(* IEC 61131-3 sources: TetherPLC/compat/tc2, 47 files *)

(* ---- tc2_math.st ---- *)
// Tc2_Math compatibility functions (TwinCAT 3 PLC Library Tc2_Math).
// Pure LREAL math; sources from docs/plc/plan/21-twincat-libraries.md §7.
// Limitation: TRUNC narrows through DINT, so |x| >= 2^31 loses precision
// (same bound as Beckhoff's 32-bit TRUNC-based implementations).

FUNCTION F_TruncL : LREAL
VAR_INPUT
    lr_in : LREAL;
END_VAR
    F_TruncL := DINT_TO_LREAL(TRUNC(lr_in));
END_FUNCTION

FUNCTION CEIL : LREAL
VAR_INPUT
    lr_in : LREAL;
END_VAR
VAR
    t : LREAL;
END_VAR
    t := F_TruncL(lr_in);
    IF lr_in > t THEN
        CEIL := t + 1.0;
    ELSE
        CEIL := t;
    END_IF;
END_FUNCTION

FUNCTION FLOOR : LREAL
VAR_INPUT
    lr_in : LREAL;
END_VAR
VAR
    t : LREAL;
END_VAR
    t := F_TruncL(lr_in);
    IF lr_in < t THEN
        FLOOR := t - 1.0;
    ELSE
        FLOOR := t;
    END_IF;
END_FUNCTION

FUNCTION FRAC : LREAL
VAR_INPUT
    lr_in : LREAL;
END_VAR
    FRAC := lr_in - F_TruncL(lr_in);
END_FUNCTION

FUNCTION LTRUNC : LREAL
VAR_INPUT
    lr_in : LREAL;
END_VAR
    LTRUNC := F_TruncL(lr_in);
END_FUNCTION

FUNCTION LMOD : LREAL
VAR_INPUT
    lr_Value : LREAL;
    lr_Arg   : LREAL;
END_VAR
    IF lr_Arg = 0.0 THEN
        LMOD := 0.0;
    ELSE
        LMOD := lr_Value - F_TruncL(lr_Value / lr_Arg) * lr_Arg;
    END_IF;
END_FUNCTION

FUNCTION MODABS : LREAL
VAR_INPUT
    lr_val : LREAL;
    lr_mod : LREAL;
END_VAR
VAR
    am : LREAL;
END_VAR
    am := ABS(lr_mod);
    IF am = 0.0 THEN
        MODABS := 0.0;
    ELSE
        MODABS := lr_val - FLOOR(lr_val / am) * am;
    END_IF;
END_FUNCTION

FUNCTION MODTURNS : DINT
VAR_INPUT
    lr_Value : LREAL;
    lr_Arg   : LREAL;
END_VAR
    IF lr_Arg = 0.0 THEN
        MODTURNS := 0;
    ELSE
        MODTURNS := TRUNC(lr_Value / lr_Arg);
    END_IF;
END_FUNCTION

FUNCTION F_GetVersionTcMath : UINT
VAR_INPUT
    nVersionElement : INT;
END_VAR
    F_GetVersionTcMath := 16#0100;
END_FUNCTION

(* ---- tc2_ncdrive.st ---- *)
// Tc2_NcDrive — NC-axis SoE/CoE drive blocks.
//
// The 20 function blocks of this library are provided by
// compat/tc2/tc2_mc2_drive.st: the NcDrive variants take
// NCTOPLC_AXIS_REF + sNetId where the MC2_Drive variants take
// AXIS_REF + NetId, and both flatten to the same UDINT axis handle
// (slave = Axis - 1) over FB_Soe/FB_MotionAxis.  Covered:
//   FB_SoEReset, FB_SoEWritePassword, FB_SoEExecuteCommand,
//   FB_SoEWriteCommandControl, FB_SoEReadCommandState,
//   FB_SoEReadDiagMessage, FB_SoEReadDiagNumber,
//   FB_SoEReadDiagNumberList, FB_SoEReadClassXDiag, FB_SoERead,
//   FB_SoEWrite, FB_SoEReadAmplifierTemperature,
//   FB_SoEReadMotorTemperature, FB_SoEReadDcBusCurrent,
//   FB_SoEReadDcBusVoltage, FB_CoERead, FB_CoEWrite,
//   FB_SoEAX5000ReadActMainVoltage, FB_SoEAX5000SetMotorCtrlWord,
//   FB_SoEAX5000FirmwareUpdate.
// Deviations (shared with Tc2_MC2_Drive): PVOID buffers flatten to
// scalar Value members, tTimeout is not modeled, bCompleteAccess is
// accepted but sub-index access is unsupported, and the AX5000
// firmware update records the request only.

// F_GetVersionTcNcDrive — library version.
FUNCTION F_GetVersionTcNcDrive : UDINT
F_GetVersionTcNcDrive := 16#0100;
END_FUNCTION

(* ---- tc2_standard_wide.st ---- *)
// Tc2_Standard wide-string functions (TwinCAT 3 PLC Library Tc2_Standard).
// W* signatures mirror IEC 61131-3 string functions; bodies delegate to the
// same builtins, which already accept WSTRING operands.
// Sources: docs/plc/plan/21-twincat-libraries.md §7.

FUNCTION WCONCAT : WSTRING
VAR_INPUT
    STR1 : WSTRING;
    STR2 : WSTRING;
END_VAR
    WCONCAT := CONCAT(STR1, STR2);
END_FUNCTION

FUNCTION WDELETE : WSTRING
VAR_INPUT
    STR1 : WSTRING;
    LEN  : INT;
    POS  : INT;
END_VAR
    WDELETE := DELETE(STR1, LEN, POS);
END_FUNCTION

FUNCTION WFIND : INT
VAR_INPUT
    STR1 : WSTRING;
    STR2 : WSTRING;
END_VAR
    WFIND := FIND(STR1, STR2);
END_FUNCTION

FUNCTION WINSERT : WSTRING
VAR_INPUT
    STR1 : WSTRING;
    STR2 : WSTRING;
    POS  : INT;
END_VAR
    WINSERT := INSERT(STR1, STR2, POS);
END_FUNCTION

FUNCTION WLEFT : WSTRING
VAR_INPUT
    STR  : WSTRING;
    SIZE : INT;
END_VAR
    WLEFT := LEFT(STR, SIZE);
END_FUNCTION

FUNCTION WLEN : INT
VAR_INPUT
    STR : WSTRING;
END_VAR
    WLEN := LEN(STR);
END_FUNCTION

FUNCTION WMID : WSTRING
VAR_INPUT
    STR  : WSTRING;
    LEN  : INT;
    POS  : INT;
END_VAR
    WMID := MID(STR, LEN, POS);
END_FUNCTION

FUNCTION WREPLACE : WSTRING
VAR_INPUT
    STR1 : WSTRING;
    STR2 : WSTRING;
    L    : INT;
    P    : INT;
END_VAR
    WREPLACE := REPLACE(STR1, STR2, L, P);
END_FUNCTION

FUNCTION WRIGHT : WSTRING
VAR_INPUT
    STR  : WSTRING;
    SIZE : INT;
END_VAR
    WRIGHT := RIGHT(STR, SIZE);
END_FUNCTION

(* ---- tc2_aes70.st ---- *)
// tc2_aes70.st — TwinCAT audio-control client surface (Tc3_AES70 /
// TF6301-ish shape) over the tplc-aes70 service + FB_Aes70 builtin.
//
// The PLC is the OCA client over OSCP TCP (AES70/Open Control
// Architecture): FB_Aes70Connect opens the TCP session on the OCA
// control port (default 65000); FB_Aes70Call carries an OcaCommand
// (targetONo + methodID + parameter bytes);
// FB_Aes70Receive polls for a pending OcaResponse each scan;
// Keepalive sends an OSCP heartbeat; Disconnect releases.
//
// Parameters and response payloads are raw bytes bounded
// STRING[255] — the caller composes/parses the OCA-serialized
// parameter set.  Notification subscriptions, the full OCA class
// catalog, and property/get-set shorthands are out of scope for
// this tranche.

// ---- FB_Aes70Connect: TCP session on the OCA control port ----
FUNCTION_BLOCK FB_Aes70Connect
VAR_INPUT
    Execute : BOOL;
    Host : STRING[63];
    Port : UDINT;
END_VAR
VAR_OUTPUT
    Done : BOOL;
    Busy : BOOL;
    Error : BOOL;
    ErrorID : UDINT;
    ConnectionHdl : UDINT;
END_VAR
VAR
    ch : FB_Aes70;
    exPrev : BOOL;
END_VAR
    Done := FALSE;
    Error := FALSE;
    ErrorID := 0;
    IF Execute AND NOT exPrev THEN
        ch.OP := 1;
        ch.HOST := Host;
        ch.PORT := Port;
        ch();
        IF ch.STATUS = 0 THEN
            Done := TRUE;
            ConnectionHdl := ch.HANDLE;
        ELSE
            Error := TRUE;
            ErrorID := ch.ERRID;
        END_IF;
    END_IF;
    exPrev := Execute;
    Busy := FALSE;
END_FUNCTION_BLOCK

// ---- FB_Aes70Disconnect: release the session ----
FUNCTION_BLOCK FB_Aes70Disconnect
VAR_INPUT
    Execute : BOOL;
    ConnectionHdl : UDINT;
END_VAR
VAR_OUTPUT
    Done : BOOL;
    Busy : BOOL;
    Error : BOOL;
    ErrorID : UDINT;
END_VAR
VAR
    ch : FB_Aes70;
    exPrev : BOOL;
END_VAR
    Done := FALSE;
    Error := FALSE;
    ErrorID := 0;
    IF Execute AND NOT exPrev THEN
        ch.OP := 2;
        ch.HANDLE := ConnectionHdl;
        ch();
        IF ch.STATUS = 0 THEN
            Done := TRUE;
        ELSE
            Error := TRUE;
            ErrorID := ch.ERRID;
        END_IF;
    END_IF;
    exPrev := Execute;
    Busy := FALSE;
END_FUNCTION_BLOCK

// ---- FB_Aes70Call: OcaCommand on an object ----
FUNCTION_BLOCK FB_Aes70Call
VAR_INPUT
    Execute : BOOL;
    ConnectionHdl : UDINT;
    TargetONo : UDINT;
    MethodID : UDINT;
    Params : STRING[255];
END_VAR
VAR_OUTPUT
    Done : BOOL;
    Error : BOOL;
    ErrorID : UDINT;
    RequestHdl : UDINT;
END_VAR
VAR
    ch : FB_Aes70;
    exPrev : BOOL;
END_VAR
    Done := FALSE;
    Error := FALSE;
    ErrorID := 0;
    IF Execute AND NOT exPrev THEN
        ch.OP := 4;
        ch.HANDLE := ConnectionHdl;
        ch.TARGET := TargetONo;
        ch.METH := MethodID;
        ch.PARAMS := Params;
        ch();
        IF ch.STATUS = 0 THEN
            Done := TRUE;
            RequestHdl := ch.HANDLE2;
        ELSE
            Error := TRUE;
            ErrorID := ch.ERRID;
        END_IF;
    END_IF;
    exPrev := Execute;
END_FUNCTION_BLOCK

// ---- FB_Aes70Keepalive: OSCP heartbeat ----
FUNCTION_BLOCK FB_Aes70Keepalive
VAR_INPUT
    Execute : BOOL;
    ConnectionHdl : UDINT;
END_VAR
VAR_OUTPUT
    Done : BOOL;
    Error : BOOL;
    ErrorID : UDINT;
END_VAR
VAR
    ch : FB_Aes70;
    exPrev : BOOL;
END_VAR
    Done := FALSE;
    Error := FALSE;
    ErrorID := 0;
    IF Execute AND NOT exPrev THEN
        ch.OP := 5;
        ch.HANDLE := ConnectionHdl;
        ch();
        IF ch.STATUS = 0 THEN
            Done := TRUE;
        ELSE
            Error := TRUE;
            ErrorID := ch.ERRID;
        END_IF;
    END_IF;
    exPrev := Execute;
END_FUNCTION_BLOCK

// ---- FB_Aes70Receive: poll for a pending OcaResponse ----
FUNCTION_BLOCK FB_Aes70Receive
VAR_INPUT
    Execute : BOOL;
    ConnectionHdl : UDINT;
END_VAR
VAR_OUTPUT
    Done : BOOL;
    Message : BOOL;
    Error : BOOL;
    ErrorID : UDINT;
    RequestHdl : UDINT;
    StatusCode : UDINT;
    Payload : STRING[255];
END_VAR
VAR
    ch : FB_Aes70;
END_VAR
    Done := FALSE;
    Message := FALSE;
    Error := FALSE;
    ErrorID := 0;
    IF Execute THEN
        ch.OP := 6;
        ch.HANDLE := ConnectionHdl;
        ch();
        IF ch.STATUS >= 0 THEN
            Done := TRUE;
            Message := TRUE;
            RequestHdl := ch.HANDLE2;
            StatusCode := ch.STATUSCODE;
            Payload := ch.RXPAYLOAD;
        ELSIF ch.STATUS = 1 THEN
            Done := TRUE;
        ELSE
            Error := TRUE;
            ErrorID := ch.ERRID;
        END_IF;
    END_IF;
END_FUNCTION_BLOCK

(* ---- tc2_babasic.st ---- *)
// tc2_babasic.st — Tc2_BABasic surface (TF8010_TC3_BABasic_EN):
// pure-ST building-automation blocks — no host/hardware
// dependency.  Covers the documented categories: conversion,
// energy management, facade, lighting, scenes, signal
// processing, and timers.  Remaining catalogue entries are
// variants of the same patterns (documented gap notes in the
// plan file).

// ---- F_Scale: linear rescale ----
FUNCTION F_Scale : LREAL
VAR_INPUT
    x : LREAL;
    xMin : LREAL;
    xMax : LREAL;
    yMin : LREAL;
    yMax : LREAL;
END_VAR
    IF xMax = xMin THEN
        F_Scale := yMin;
    ELSE
        F_Scale := yMin + (x - xMin) * (yMax - yMin) / (xMax - xMin);
    END_IF;
END_FUNCTION

// ---- FB_ThresholdSwitch: two-point switch with hysteresis ----
FUNCTION_BLOCK FB_ThresholdSwitch
VAR_INPUT
    x : LREAL;
    On : LREAL;                 // switch on when x >= On
    Off : LREAL;                // switch off when x <= Off
END_VAR
VAR_OUTPUT
    Q : BOOL;
END_VAR
    IF x >= On THEN Q := TRUE; END_IF;
    IF x <= Off THEN Q := FALSE; END_IF;
END_FUNCTION_BLOCK

// ---- FB_ShortLongClick: click length discrimination ----
// A release before tLong reports Short; holding past tLong
// reports Long.
FUNCTION_BLOCK FB_ShortLongClick
VAR_INPUT
    In : BOOL;
    tLong : LREAL;              // s
    CycleTime : LREAL;          // s
END_VAR
VAR_OUTPUT
    Short : BOOL;
    Long : BOOL;
END_VAR
VAR
    tAcc : LREAL;
    prev : BOOL;
END_VAR
    Short := FALSE;
    Long := FALSE;
    IF CycleTime <= 0.0 THEN RETURN; END_IF;
    IF In THEN
        tAcc := tAcc + CycleTime;
        IF tAcc >= tLong AND NOT prev THEN
            Long := TRUE;      // edge: just passed threshold
        END_IF;
    ELSE
        IF tAcc > 0.0 AND tAcc < tLong THEN
            Short := TRUE;     // released early
        END_IF;
        tAcc := 0.0;
    END_IF;
    prev := tAcc >= tLong;
END_FUNCTION_BLOCK

// ---- FB_SingleDoubleClick: single vs double click ----
FUNCTION_BLOCK FB_SingleDoubleClick
VAR_INPUT
    In : BOOL;
    tDouble : LREAL;            // s window for second click
    CycleTime : LREAL;
END_VAR
VAR_OUTPUT
    Single : BOOL;
    Double : BOOL;
END_VAR
VAR
    clicks : INT;
    tGap : LREAL;
    prev : BOOL;
END_VAR
    Single := FALSE;
    Double := FALSE;
    IF CycleTime <= 0.0 THEN RETURN; END_IF;
    IF In AND NOT prev THEN
        clicks := clicks + 1;
    END_IF;
    prev := In;
    IF clicks > 0 AND NOT In THEN
        tGap := tGap + CycleTime;
        IF tGap >= tDouble THEN
            IF clicks = 1 THEN
                Single := TRUE;
            ELSE
                Double := TRUE;
            END_IF;
            clicks := 0;
            tGap := 0.0;
        END_IF;
    ELSIF In THEN
        tGap := 0.0;
    END_IF;
END_FUNCTION_BLOCK

// ---- FB_SignallingContact: latch until acknowledged ----
FUNCTION_BLOCK FB_SignallingContact
VAR_INPUT
    In : BOOL;
    Ack : BOOL;
END_VAR
VAR_OUTPUT
    Q : BOOL;
END_VAR
    IF In THEN Q := TRUE; END_IF;
    IF Ack THEN Q := FALSE; END_IF;
END_FUNCTION_BLOCK

// ---- FB_Ramp: slew-rate limiter ----
FUNCTION_BLOCK FB_Ramp
VAR_INPUT
    Enable : BOOL;
    Setpoint : LREAL;
    SlewUp : LREAL;             // unit/s
    SlewDown : LREAL;
    CycleTime : LREAL;
END_VAR
VAR_OUTPUT
    Out : LREAL;
    AtTarget : BOOL;
END_VAR
    IF NOT Enable THEN
        AtTarget := FALSE;
        RETURN;
    END_IF;
    IF Out < Setpoint THEN
        Out := Out + SlewUp * CycleTime;
        IF Out > Setpoint THEN Out := Setpoint; END_IF;
    ELSIF Out > Setpoint THEN
        Out := Out - SlewDown * CycleTime;
        IF Out < Setpoint THEN Out := Setpoint; END_IF;
    END_IF;
    AtTarget := Out = Setpoint;
END_FUNCTION_BLOCK

// ---- FB_Light: light channel with off-delay ----
FUNCTION_BLOCK FB_Light
VAR_INPUT
    On : BOOL;
    OffDelay : LREAL;           // s; 0 = no delay
    CycleTime : LREAL;
END_VAR
VAR_OUTPUT
    Q : BOOL;
    TimeLeft : LREAL;
END_VAR
VAR
    tLeft : LREAL;
END_VAR
    IF On THEN
        tLeft := OffDelay;
        Q := TRUE;
    ELSIF tLeft > 0.0 THEN
        tLeft := tLeft - CycleTime;
        Q := tLeft > 0.0;
    ELSE
        Q := FALSE;
    END_IF;
    TimeLeft := tLeft;
END_FUNCTION_BLOCK

// ---- FB_StairwellLight: retriggable stairwell timer ----
FUNCTION_BLOCK FB_StairwellLight
VAR_INPUT
    Trigger : BOOL;
    Duration : LREAL;           // s
    CycleTime : LREAL;
END_VAR
VAR_OUTPUT
    Q : BOOL;
    TimeLeft : LREAL;
END_VAR
VAR
    tLeft : LREAL;
END_VAR
    IF Trigger THEN tLeft := Duration; END_IF;
    IF tLeft > 0.0 THEN
        tLeft := tLeft - CycleTime;
        Q := TRUE;
    ELSE
        tLeft := 0.0;
        Q := FALSE;
    END_IF;
    TimeLeft := tLeft;
END_FUNCTION_BLOCK

// ---- FB_Dimmer1Switch: one-button dimmer ----
// Short click toggles on/off (memory of last level); long press
// ramps the level between Lo and Hi.
FUNCTION_BLOCK FB_Dimmer1Switch
VAR_INPUT
    Click : FB_ShortLongClick;
    LevelHi : LREAL;            // max level (e.g. 100)
    LevelLo : LREAL;
    SlewRate : LREAL;           // level/s
    CycleTime : LREAL;
END_VAR
VAR_OUTPUT
    Level : LREAL;
    Q : BOOL;
END_VAR
VAR
    mem : LREAL;
    dir : INT;
    ramp : FB_Ramp;
END_VAR
    Click();
    IF Click.Short THEN
        IF Q THEN
            mem := Level;
            Q := FALSE;
        ELSE
            Q := TRUE;
        END_IF;
    END_IF;
    IF Click.Long THEN dir := -dir; END_IF;
    ramp.Enable := TRUE;
    IF Q THEN
        IF dir = 0 THEN dir := 1; END_IF;
        IF Click.In THEN
            IF dir > 0 THEN
                ramp.Setpoint := LevelHi;
            ELSE
                ramp.Setpoint := LevelLo;
            END_IF;
        ELSE
            ramp.Setpoint := LevelHi;
        END_IF;
    ELSE
        ramp.Setpoint := 0.0;
    END_IF;
    ramp.SlewUp := SlewRate;
    ramp.SlewDown := SlewRate;
    ramp.CycleTime := CycleTime;
    ramp();
    Level := ramp.Out;
END_FUNCTION_BLOCK

// ---- FB_Dimmer2Switch: two-button up/down dimmer ----
// bUp/bDown short: on at max / off.  Long: ramp while held.
FUNCTION_BLOCK FB_Dimmer2Switch
VAR_INPUT
    bUp : BOOL;
    bDown : BOOL;
    LevelHi : LREAL;
    LevelLo : LREAL;
    SlewRate : LREAL;
    tLong : LREAL;
    CycleTime : LREAL;
END_VAR
VAR_OUTPUT
    Level : LREAL;
    Q : BOOL;
END_VAR
VAR
    tUp : LREAL;
    tDown : LREAL;
    upP : BOOL;
    downP : BOOL;
END_VAR
    IF bUp THEN tUp := tUp + CycleTime; ELSE tUp := 0.0; END_IF;
    IF bDown THEN tDown := tDown + CycleTime; ELSE tDown := 0.0; END_IF;
    // short-click edges on release
    IF NOT bUp AND upP AND tUp > 0.0 AND tUp < tLong THEN
        Q := TRUE; Level := LevelHi;
    END_IF;
    IF NOT bDown AND downP AND tDown > 0.0 AND tDown < tLong THEN
        Q := FALSE; Level := 0.0;
    END_IF;
    // long-press ramp
    IF tUp >= tLong THEN
        Level := Level + SlewRate * CycleTime;
        IF Level > LevelHi THEN Level := LevelHi; END_IF;
        Q := TRUE;
    END_IF;
    IF tDown >= tLong THEN
        Level := Level - SlewRate * CycleTime;
        IF Level < 0.0 THEN Level := 0.0; END_IF;
        IF Level <= LevelLo THEN Q := FALSE; END_IF;
    END_IF;
    upP := bUp;
    downP := bDown;
END_FUNCTION_BLOCK

// ---- FB_VenetianBlind: blind with slat-angle control ----
// up/down drive position (0 = open/top, PosMax = closed);
// a short tap nudges the slat angle instead.
FUNCTION_BLOCK FB_VenetianBlind
VAR_INPUT
    bUp : BOOL;
    bDown : BOOL;
    PosMax : LREAL;             // s travel top->bottom
    SlatMax : LREAL;            // s slat full swing
    tSlat : LREAL;              // tap threshold
    CycleTime : LREAL;
END_VAR
VAR_OUTPUT
    Position : LREAL;           // 0..PosMax
    Slat : LREAL;               // -SlatMax..+SlatMax
END_VAR
VAR
    tDir : LREAL;
    upP : BOOL;
    downP : BOOL;
END_VAR
    IF bUp THEN
        tDir := tDir + CycleTime;
        IF tDir >= tSlat THEN
            Position := Position - CycleTime;
            IF Position < 0.0 THEN Position := 0.0; END_IF;
        END_IF;
    END_IF;
    IF bDown THEN
        tDir := tDir + CycleTime;
        IF tDir >= tSlat THEN
            Position := Position + CycleTime;
            IF Position > PosMax THEN Position := PosMax; END_IF;
        END_IF;
    END_IF;
    // released early: slat nudge in that direction
    IF NOT bUp AND upP AND tDir > 0.0 AND tDir < tSlat THEN
        Slat := Slat - CycleTime * 4.0;
        IF Slat < -SlatMax THEN Slat := -SlatMax; END_IF;
    END_IF;
    IF NOT bDown AND downP AND tDir > 0.0 AND tDir < tSlat THEN
        Slat := Slat + CycleTime * 4.0;
        IF Slat > SlatMax THEN Slat := SlatMax; END_IF;
    END_IF;
    IF NOT bUp AND NOT bDown THEN tDir := 0.0; END_IF;
    upP := bUp;
    downP := bDown;
END_FUNCTION_BLOCK

// ---- FB_MaximumDemandController: shed loads over limit ----
// Counts active inputs; when the count exceeds Limit, outputs
// are shed starting from the highest index (shed mask).
FUNCTION_BLOCK FB_MaximumDemandController
VAR_INPUT
    In1 : BOOL;
    In2 : BOOL;
    In3 : BOOL;
    In4 : BOOL;
    Limit : INT;
    Enable : BOOL;
END_VAR
VAR_OUTPUT
    Q1 : BOOL;
    Q2 : BOOL;
    Q3 : BOOL;
    Q4 : BOOL;
    Shedding : BOOL;
    Active : INT;
END_VAR
VAR
    n : INT;
END_VAR
    IF NOT Enable THEN
        Q1 := FALSE; Q2 := FALSE; Q3 := FALSE; Q4 := FALSE;
        Shedding := FALSE;
        Active := 0;
        RETURN;
    END_IF;
    n := 0;
    IF In1 THEN n := n + 1; END_IF;
    IF In2 THEN n := n + 1; END_IF;
    IF In3 THEN n := n + 1; END_IF;
    IF In4 THEN n := n + 1; END_IF;
    Active := n;
    Q1 := In1; Q2 := In2; Q3 := In3; Q4 := In4;
    Shedding := FALSE;
    IF n > Limit THEN
        Shedding := TRUE;
        // shed highest first until under limit
        IF Q4 AND n > Limit THEN Q4 := FALSE; n := n - 1; END_IF;
        IF Q3 AND n > Limit THEN Q3 := FALSE; n := n - 1; END_IF;
        IF Q2 AND n > Limit THEN Q2 := FALSE; n := n - 1; END_IF;
        IF Q1 AND n > Limit THEN Q1 := FALSE; n := n - 1; END_IF;
    END_IF;
END_FUNCTION_BLOCK

// ---- FB_DailyScheduler: on/off windows within a day ----
// MinuteOfDay 0..1439; on when inside [OnMin, OffMin).
FUNCTION_BLOCK FB_DailyScheduler
VAR_INPUT
    MinuteOfDay : INT;
    OnMin : INT;
    OffMin : INT;
    Enable : BOOL;
END_VAR
VAR_OUTPUT
    Q : BOOL;
END_VAR
    IF NOT Enable THEN Q := FALSE; RETURN; END_IF;
    IF OnMin < OffMin THEN
        Q := MinuteOfDay >= OnMin AND MinuteOfDay < OffMin;
    ELSE
        // window wraps midnight
        Q := MinuteOfDay >= OnMin OR MinuteOfDay < OffMin;
    END_IF;
END_FUNCTION_BLOCK

// ---- FB_ScenesLighting: recall one of N light levels ----
FUNCTION_BLOCK FB_ScenesLighting
VAR_INPUT
    Scene : INT;                // 1..4
    L1 : LREAL;
    L2 : LREAL;
    L3 : LREAL;
    L4 : LREAL;
    Enable : BOOL;
END_VAR
VAR_OUTPUT
    Level : LREAL;
    Q : BOOL;
END_VAR
    IF NOT Enable THEN
        Level := 0.0; Q := FALSE;
        RETURN;
    END_IF;
    IF Scene = 1 THEN Level := L1;
    ELSIF Scene = 2 THEN Level := L2;
    ELSIF Scene = 3 THEN Level := L3;
    ELSIF Scene = 4 THEN Level := L4;
    ELSE Level := 0.0;
    END_IF;
    Q := Level > 0.0;
END_FUNCTION_BLOCK

(* ---- tc2_cm.st ---- *)
// tc2_cm.st — Tc2_CM (curve/math) surface — curve and math
// primitives, pure-ST, no service or hardware.
//
// These are the curve/trajectory helpers: a function generator
// (sawtooth/triangle/square), a piecewise-linear interpolator over
// a breakpoint table, and a cam-style master->slave curve
// (linear segment lookup between master positions).  All take
// phase/cycle inputs from the caller.

// ---- FB_FuncGen: periodic function generator ----
// Shape: 0=sawtooth, 1=triangle, 2=square
FUNCTION_BLOCK FB_FuncGen
VAR_INPUT
    Execute : BOOL;
    Shape : UDINT;          // 0=saw 1=tri 2=square
    Period : LREAL;         // period (s), >0
    Amplitude : LREAL;
    Offset : LREAL;
    CycleTime : LREAL;
END_VAR
VAR_OUTPUT
    Done : BOOL;
    Output : LREAL;
    Phase : LREAL;          // 0..1
END_VAR
VAR
    ph : LREAL;
    y : LREAL;
END_VAR
    Done := FALSE;
    IF Execute AND Period > 0.0 THEN
        ph := ph + CycleTime / Period;
        IF ph >= 1.0 THEN ph := ph - 1.0; END_IF;
        IF Shape = 0 THEN
            y := ph;                                   // sawtooth
        ELSIF Shape = 1 THEN
            IF ph < 0.5 THEN
                y := 2.0 * ph;                          // triangle up
            ELSE
                y := 2.0 * (1.0 - ph);                  // triangle down
            END_IF;
        ELSE
            IF ph < 0.5 THEN
                y := 1.0;                               // square high
            ELSE
                y := 0.0;                               // square low
            END_IF;
        END_IF;
        Output := Offset + Amplitude * y;
        Phase := ph;
        Done := TRUE;
    END_IF;
END_FUNCTION_BLOCK

// ---- FB_LinInterp: piecewise-linear interpolation over a table ----
// PointsX[i] -> PointsY[i], clamped at the ends.  Caller fills the
// 8-point table.
FUNCTION_BLOCK FB_LinInterp
VAR_INPUT
    Execute : BOOL;
    X : LREAL;
    X0 : LREAL; Y0 : LREAL;
    X1 : LREAL; Y1 : LREAL;
    X2 : LREAL; Y2 : LREAL;
    X3 : LREAL; Y3 : LREAL;
END_VAR
VAR_OUTPUT
    Done : BOOL;
    Error : BOOL;
    ErrorID : UDINT;
    Y : LREAL;
END_VAR
    Done := FALSE;
    Error := FALSE;
    ErrorID := 0;
    IF NOT Execute THEN RETURN; END_IF;
    // 4-point piecewise-linear — X0..X3 ascending
    IF X <= X1 THEN
        IF X1 = X0 THEN Error := TRUE; ErrorID := 1; END_IF;
        Y := Y0 + (Y1 - Y0) * (X - X0) / (X1 - X0);
    ELSIF X <= X2 THEN
        IF X2 = X1 THEN Error := TRUE; ErrorID := 1; END_IF;
        Y := Y1 + (Y2 - Y1) * (X - X1) / (X2 - X1);
    ELSIF X <= X3 THEN
        IF X3 = X2 THEN Error := TRUE; ErrorID := 1; END_IF;
        Y := Y2 + (Y3 - Y2) * (X - X2) / (X3 - X2);
    ELSE
        Y := Y3;   // clamp above
    END_IF;
    IF NOT Error THEN Done := TRUE; END_IF;
END_FUNCTION_BLOCK

// ---- FB_CamProfile: master-position -> slave-position cam ----
// A simple linear cam: slave ramps 0..SlaveAmp as master goes
// 0..MasterEnd, then holds.  Model for a cam table lookup.
FUNCTION_BLOCK FB_CamProfile
VAR_INPUT
    Execute : BOOL;
    Master : LREAL;         // master position
    MasterEnd : LREAL;      // master end (cam period), >0
    SlaveAmp : LREAL;       // slave amplitude
END_VAR
VAR_OUTPUT
    Done : BOOL;
    Slave : LREAL;
    InSync : BOOL;
END_VAR
VAR
    k : LREAL;
END_VAR
    Done := FALSE;
    IF Execute AND MasterEnd > 0.0 THEN
        k := Master;
        IF k < 0.0 THEN k := 0.0; END_IF;
        IF k > MasterEnd THEN k := MasterEnd; END_IF;
        Slave := SlaveAmp * k / MasterEnd;
        InSync := (Master >= 0.0) AND (Master <= MasterEnd);
        Done := TRUE;
    END_IF;
END_FUNCTION_BLOCK

(* ---- tc2_controllertoolbox.st ---- *)
// tc2_controllertoolbox.st — Tc2_ControllerToolbox surface —
// additional controller primitives, pure-ST, no service or
// hardware: dead-time delay, hysteresis / two-position /
// three-position controllers, PWM duty converter, and
// running statistics (mean + standard deviation).
//
// All blocks take CycleTime as a VAR_INPUT (the caller's scan
// period, TwinCAT's T_PLC_US pattern).  DeadTime holds a ring of
// samples and outputs the N-cycle-delayed value.

// ---- FB_DeadTime: delay a signal N cycles ----
FUNCTION_BLOCK FB_DeadTime
VAR_INPUT
    Execute : BOOL;
    Input : LREAL;
    DelayCycles : UDINT;   // 0..63
END_VAR
VAR_OUTPUT
    Done : BOOL;
    Output : LREAL;
END_VAR
VAR
    buf : ARRAY[0..63] OF LREAL;
    idx : UDINT;
END_VAR
    Done := FALSE;
    IF Execute THEN
        buf[idx] := Input;
        Output := buf[(idx + 64 - (DelayCycles MOD 64)) MOD 64];
        idx := (idx + 1) MOD 64;
        Done := TRUE;
    END_IF;
END_FUNCTION_BLOCK

// ---- FB_Hysteresis: relay with on/off hysteresis band ----
FUNCTION_BLOCK FB_Hysteresis
VAR_INPUT
    Execute : BOOL;
    Input : LREAL;
    OnLevel : LREAL;   // switch ON at/below
    OffLevel : LREAL;  // switch OFF at/above (Off > On)
END_VAR
VAR_OUTPUT
    Done : BOOL;
    Out : BOOL;
END_VAR
VAR
    on : BOOL;
END_VAR
    Done := FALSE;
    IF Execute THEN
        IF Input <= OnLevel THEN
            on := TRUE;
        ELSIF Input >= OffLevel THEN
            on := FALSE;
        END_IF;
        Out := on;
        Done := TRUE;
    END_IF;
END_FUNCTION_BLOCK

// ---- FB_TwoPosition: two-position (on/off) controller ----
FUNCTION_BLOCK FB_TwoPosition
VAR_INPUT
    Execute : BOOL;
    Setpoint : LREAL;
    Actual : LREAL;
    Hysteresis : LREAL;   // +- band around Setpoint
END_VAR
VAR_OUTPUT
    Done : BOOL;
    Out : BOOL;           // TRUE = drive high
END_VAR
VAR
    e : LREAL;
END_VAR
    Done := FALSE;
    IF Execute THEN
        e := Setpoint - Actual;
        IF e > Hysteresis THEN
            Out := TRUE;      // below band -> drive on
        ELSIF e < -Hysteresis THEN
            Out := FALSE;     // above band -> drive off
        END_IF;
        Done := TRUE;
    END_IF;
END_FUNCTION_BLOCK

// ---- FB_ThreePosition: three-position controller ----
FUNCTION_BLOCK FB_ThreePosition
VAR_INPUT
    Execute : BOOL;
    Setpoint : LREAL;
    Actual : LREAL;
    Deadband : LREAL;     // +- neutral zone
    Hysteresis : LREAL;   // +- switch band beyond deadband
END_VAR
VAR_OUTPUT
    Done : BOOL;
    OutPos : INT;         // -1 = low, 0 = neutral, +1 = high
END_VAR
VAR
    e : LREAL;
END_VAR
    Done := FALSE;
    IF Execute THEN
        e := Setpoint - Actual;
        IF e > Deadband + Hysteresis THEN
            OutPos := 1;      // well below -> drive high
        ELSIF e < -Deadband - Hysteresis THEN
            OutPos := -1;     // well above -> drive low
        ELSIF e > -Deadband AND e < Deadband THEN
            OutPos := 0;      // inside deadband -> neutral
        END_IF;
        // else keep prior OutPos (hysteresis band)
        Done := TRUE;
    END_IF;
END_FUNCTION_BLOCK

// ---- FB_Statistics: running mean + standard deviation ----
FUNCTION_BLOCK FB_Statistics
VAR_INPUT
    Execute : BOOL;
    Input : LREAL;
    N : UDINT;            // 1..64 — window length
END_VAR
VAR_OUTPUT
    Done : BOOL;
    Mean : LREAL;
    StdDev : LREAL;
    Minimum : LREAL;
    Maximum : LREAL;
END_VAR
VAR
    buf : ARRAY[0..63] OF LREAL;
    idx : UDINT;
    cnt : UDINT;
    i : UDINT;
    s : LREAL;
    v : LREAL;
    m : LREAL;
    lo : LREAL;
    hi : LREAL;
    nR : LREAL;
    x : LREAL;     // Newton's sqrt iterate
    it : UDINT;
END_VAR
    Done := FALSE;
    IF Execute AND N > 0 AND N <= 64 THEN
        buf[idx] := Input;
        idx := (idx + 1);
        IF idx >= N THEN idx := 0; END_IF;
        IF cnt < N THEN cnt := cnt + 1; END_IF;
        s := 0.0; lo := buf[0]; hi := buf[0];
        FOR i := 0 TO 63 BY 1 DO
            IF i < cnt THEN
                s := s + buf[i];
                IF buf[i] < lo THEN lo := buf[i]; END_IF;
                IF buf[i] > hi THEN hi := buf[i]; END_IF;
            END_IF;
        END_FOR;
        nR := DINT_TO_LREAL(UDINT_TO_DINT(cnt));
        m := s / nR;
        v := 0.0;
        FOR i := 0 TO 63 BY 1 DO
            IF i < cnt THEN
                v := v + (buf[i] - m) * (buf[i] - m);
            END_IF;
        END_FOR;
        v := v / nR;
        // StdDev = sqrt(v) via Newton's method — no SQRT builtin
        IF v <= 0.0 THEN
            StdDev := 0.0;
        ELSE
            x := v;
            FOR it := 1 TO 12 BY 1 DO
                x := 0.5 * (x + v / x);
            END_FOR;
            StdDev := x;
        END_IF;
        Mean := m;
        Minimum := lo;
        Maximum := hi;
        Done := TRUE;
    END_IF;
END_FUNCTION_BLOCK

// ---- FB_Pwm: duty-cycle converter (0..100% -> pulse width) ----
FUNCTION_BLOCK FB_Pwm
VAR_INPUT
    Execute : BOOL;
    Duty : LREAL;         // 0..100 percent
    Period : LREAL;       // period (s), >0
    CycleTime : LREAL;
END_VAR
VAR_OUTPUT
    Done : BOOL;
    Out : BOOL;           // TRUE during on-phase
END_VAR
VAR
    t : LREAL;            // phase accumulator (s)
    d : LREAL;
END_VAR
    Done := FALSE;
    IF Execute AND Period > 0.0 THEN
        t := t + CycleTime;
        IF t >= Period THEN t := t - Period; END_IF;
        d := Duty;
        IF d < 0.0 THEN d := 0.0; END_IF;
        IF d > 100.0 THEN d := 100.0; END_IF;
        Out := (t < Period * d / 100.0);
        Done := TRUE;
    END_IF;
END_FUNCTION_BLOCK

(* ---- tc2_dataexchange.st ---- *)
// Tc2_DataExchange -> symbolic read/write by variable name over
// the tplc-sym service (package var table -> live state blob).
// Documented differences vs. the Beckhoff library:
//   - Names address variables of the *local* program (no AMS
//     NetID routing): sNetId is accepted and ignored.
//   - Values cross typed (BOOL/DINT/LREAL): the builtin encodes
//     them into the variable's own width/type.  Byte-level access
//     is available through FB_Sym OP 1/2 for callers that need it.
//   - OnDelta blocks compare against the last transmitted value
//     and only transmit when the variable actually changed.
//   - Watchdog blocks read/write the runtime's cycle counters via
//     the same by-name path (documented reduction).

// ---- FB_ReadAdsSymByName: read a variable by name ----
FUNCTION_BLOCK FB_ReadAdsSymByName
VAR_INPUT
    bRead : BOOL;
    sNetId : STRING[23];
    sVarName : STRING[63];
END_VAR
VAR_OUTPUT
    nIntValue : DINT;
    fRealValue : LREAL;
    bBoolValue : BOOL;
    nTypeCode : UDINT;          // TPLC_IOT_* of the variable
    nSize : UDINT;              // variable size in bytes
    bBusy : BOOL;
    bError : BOOL;
    nErrorId : UDINT;
END_VAR
VAR
    sym : FB_Sym;
    prev : BOOL;
END_VAR
    bBusy := FALSE; bError := FALSE; nErrorId := 0;
    IF bRead AND NOT prev THEN
        bBusy := TRUE;
        sym.OP := 9; sym.NAME := sVarName;
        sym();
        IF sym.STATUS = 0 THEN
            IF sym.VTYP = 0 THEN
                sym.OP := 8;
            ELSIF sym.VTYP = 9 OR sym.VTYP = 10 THEN
                sym.OP := 7;
            ELSE
                sym.OP := 6;
            END_IF;
            sym();
        END_IF;
        bBusy := FALSE;
        IF sym.STATUS = 0 THEN
            nTypeCode := sym.VTYP;
            nSize := sym.SIZE;
            IF sym.VTYP = 0 THEN
                bBoolValue := sym.BB;
            ELSIF sym.VTYP = 9 OR sym.VTYP = 10 THEN
                fRealValue := sym.FB;
            ELSE
                nIntValue := sym.IB;
            END_IF;
        ELSE
            bError := TRUE; nErrorId := sym.ERRID;
        END_IF;
    END_IF;
    prev := bRead;
END_FUNCTION_BLOCK

// ---- FB_WriteAdsSymByName: write a variable by name ----
FUNCTION_BLOCK FB_WriteAdsSymByName
VAR_INPUT
    bWrite : BOOL;
    sNetId : STRING[23];
    sVarName : STRING[63];
    nIntValue : DINT;
    fRealValue : LREAL;
    bBoolValue : BOOL;
END_VAR
VAR_OUTPUT
    bBusy : BOOL;
    bDone : BOOL;
    bError : BOOL;
    nErrorId : UDINT;
END_VAR
VAR
    sym : FB_Sym;
    prev : BOOL;
END_VAR
    bBusy := FALSE; bError := FALSE; bDone := FALSE; nErrorId := 0;
    IF bWrite AND NOT prev THEN
        bBusy := TRUE;
        sym.OP := 9; sym.NAME := sVarName;
        sym();
        IF sym.STATUS = 0 THEN
            sym.IB := nIntValue; sym.FB := fRealValue; sym.BB := bBoolValue;
            IF sym.VTYP = 0 THEN
                sym.OP := 5;
            ELSIF sym.VTYP = 9 OR sym.VTYP = 10 THEN
                sym.OP := 4;
            ELSE
                sym.OP := 3;
            END_IF;
            sym();
        END_IF;
        bBusy := FALSE;
        IF sym.STATUS = 0 THEN
            bDone := TRUE;
        ELSE
            bError := TRUE; nErrorId := sym.ERRID;
        END_IF;
    END_IF;
    prev := bWrite;
END_FUNCTION_BLOCK

// ---- OnDelta writers: transmit only when the value changed ----
// One shared body per type; the delta test compares the current
// bytes against the last transmitted snapshot.
FUNCTION_BLOCK FB_WriteBoolOnDelta
VAR_INPUT
    bEnable : BOOL;
    sNetId : STRING[23];
    sVarName : STRING[63];
    bValue : BOOL;
END_VAR
VAR_OUTPUT
    bBusy : BOOL;
    bLastSignal : BOOL;
    bError : BOOL;
    nErrorId : UDINT;
    nErrorCnt : UDINT;
END_VAR
VAR
    wr : FB_WriteAdsSymByName;
    sent : BOOL;
    haveSent : BOOL;
END_VAR
    bBusy := FALSE; bError := FALSE;
    IF bEnable AND (NOT haveSent OR bValue <> sent) THEN
        bBusy := TRUE;
        wr.sVarName := sVarName;
        wr.bBoolValue := bValue;
        wr.bWrite := TRUE;
        wr();
        wr.bWrite := FALSE;
        bBusy := FALSE;
        IF wr.bError THEN
            bError := TRUE; nErrorId := wr.nErrorId;
            nErrorCnt := nErrorCnt + 1;
        ELSE
            sent := bValue; haveSent := TRUE;
            bLastSignal := bValue;
        END_IF;
    END_IF;
END_FUNCTION_BLOCK

FUNCTION_BLOCK FB_WriteByteOnDelta
VAR_INPUT
    bEnable : BOOL;
    sNetId : STRING[23];
    sVarName : STRING[63];
    nValue : BYTE;
END_VAR
VAR_OUTPUT
    bBusy : BOOL;
    nLastSignal : BYTE;
    bError : BOOL;
    nErrorId : UDINT;
    nErrorCnt : UDINT;
END_VAR
VAR
    wr : FB_WriteAdsSymByName;
    sent : BYTE;
    haveSent : BOOL;
END_VAR
    bBusy := FALSE; bError := FALSE;
    IF bEnable AND (NOT haveSent OR nValue <> sent) THEN
        bBusy := TRUE;
        wr.sVarName := sVarName;
        wr.nIntValue := BYTE_TO_DINT(nValue);
        wr.bWrite := TRUE;
        wr();
        wr.bWrite := FALSE;
        bBusy := FALSE;
        IF wr.bError THEN
            bError := TRUE; nErrorId := wr.nErrorId;
            nErrorCnt := nErrorCnt + 1;
        ELSE
            sent := nValue; haveSent := TRUE;
            nLastSignal := nValue;
        END_IF;
    END_IF;
END_FUNCTION_BLOCK

FUNCTION_BLOCK FB_WriteWordOnDelta
VAR_INPUT
    bEnable : BOOL;
    sNetId : STRING[23];
    sVarName : STRING[63];
    nValue : WORD;
END_VAR
VAR_OUTPUT
    bBusy : BOOL;
    nLastSignal : WORD;
    bError : BOOL;
    nErrorId : UDINT;
    nErrorCnt : UDINT;
END_VAR
VAR
    wr : FB_WriteAdsSymByName;
    sent : WORD;
    haveSent : BOOL;
END_VAR
    bBusy := FALSE; bError := FALSE;
    IF bEnable AND (NOT haveSent OR nValue <> sent) THEN
        bBusy := TRUE;
        wr.sVarName := sVarName;
        wr.nIntValue := WORD_TO_DINT(nValue);
        wr.bWrite := TRUE;
        wr();
        wr.bWrite := FALSE;
        bBusy := FALSE;
        IF wr.bError THEN
            bError := TRUE; nErrorId := wr.nErrorId;
            nErrorCnt := nErrorCnt + 1;
        ELSE
            sent := nValue; haveSent := TRUE;
            nLastSignal := nValue;
        END_IF;
    END_IF;
END_FUNCTION_BLOCK

FUNCTION_BLOCK FB_WriteDWordOnDelta
VAR_INPUT
    bEnable : BOOL;
    sNetId : STRING[23];
    sVarName : STRING[63];
    nValue : DWORD;
END_VAR
VAR_OUTPUT
    bBusy : BOOL;
    nLastSignal : DWORD;
    bError : BOOL;
    nErrorId : UDINT;
    nErrorCnt : UDINT;
END_VAR
VAR
    wr : FB_WriteAdsSymByName;
    sent : DWORD;
    haveSent : BOOL;
END_VAR
    bBusy := FALSE; bError := FALSE;
    IF bEnable AND (NOT haveSent OR nValue <> sent) THEN
        bBusy := TRUE;
        wr.sVarName := sVarName;
        wr.nIntValue := DWORD_TO_DINT(nValue);
        wr.bWrite := TRUE;
        wr();
        wr.bWrite := FALSE;
        bBusy := FALSE;
        IF wr.bError THEN
            bError := TRUE; nErrorId := wr.nErrorId;
            nErrorCnt := nErrorCnt + 1;
        ELSE
            sent := nValue; haveSent := TRUE;
            nLastSignal := nValue;
        END_IF;
    END_IF;
END_FUNCTION_BLOCK

FUNCTION_BLOCK FB_WriteRealOnDelta
VAR_INPUT
    bEnable : BOOL;
    sNetId : STRING[23];
    sVarName : STRING[63];
    fValue : REAL;
END_VAR
VAR_OUTPUT
    bBusy : BOOL;
    fLastSignal : REAL;
    bError : BOOL;
    nErrorId : UDINT;
    nErrorCnt : UDINT;
END_VAR
VAR
    wr : FB_WriteAdsSymByName;
    sent : REAL;
    haveSent : BOOL;
END_VAR
    bBusy := FALSE; bError := FALSE;
    IF bEnable AND (NOT haveSent OR fValue <> sent) THEN
        bBusy := TRUE;
        wr.sVarName := sVarName;
        wr.fRealValue := fValue;
        wr.bWrite := TRUE;
        wr();
        wr.bWrite := FALSE;
        bBusy := FALSE;
        IF wr.bError THEN
            bError := TRUE; nErrorId := wr.nErrorId;
            nErrorCnt := nErrorCnt + 1;
        ELSE
            sent := fValue; haveSent := TRUE;
            fLastSignal := fValue;
        END_IF;
    END_IF;
END_FUNCTION_BLOCK

FUNCTION_BLOCK FB_WriteLRealOnDelta
VAR_INPUT
    bEnable : BOOL;
    sNetId : STRING[23];
    sVarName : STRING[63];
    fValue : LREAL;
END_VAR
VAR_OUTPUT
    bBusy : BOOL;
    fLastSignal : LREAL;
    bError : BOOL;
    nErrorId : UDINT;
    nErrorCnt : UDINT;
END_VAR
VAR
    wr : FB_WriteAdsSymByName;
    sent : LREAL;
    haveSent : BOOL;
END_VAR
    bBusy := FALSE; bError := FALSE;
    IF bEnable AND (NOT haveSent OR fValue <> sent) THEN
        bBusy := TRUE;
        wr.sVarName := sVarName;
        wr.fRealValue := fValue;
        wr.bWrite := TRUE;
        wr();
        wr.bWrite := FALSE;
        bBusy := FALSE;
        IF wr.bError THEN
            bError := TRUE; nErrorId := wr.nErrorId;
            nErrorCnt := nErrorCnt + 1;
        ELSE
            sent := fValue; haveSent := TRUE;
            fLastSignal := fValue;
        END_IF;
    END_IF;
END_FUNCTION_BLOCK

// ---- Watchdog blocks ----
// FB_WriteWatchdog stamps a by-name counter variable (typically the
// program's own heartbeat), FB_CheckWatchdog verifies that a peer's
// stamp is still advancing within a timeout.
FUNCTION_BLOCK FB_WriteWatchdog
VAR_INPUT
    bEnable : BOOL;
    sNetId : STRING[23];
    sVarName : STRING[63];
END_VAR
VAR_OUTPUT
    bBusy : BOOL;
    bError : BOOL;
    nErrorId : UDINT;
    nStamps : UDINT;
END_VAR
VAR
    wr : FB_WriteAdsSymByName;
    n : DWORD;
END_VAR
    bBusy := FALSE; bError := FALSE;
    IF bEnable THEN
        n := n + 1;
        wr.sVarName := sVarName;
        wr.nIntValue := DWORD_TO_DINT(n);
        wr.bWrite := TRUE;
        wr();
        wr.bWrite := FALSE;
        IF wr.bError THEN
            bError := TRUE; nErrorId := wr.nErrorId;
        ELSE
            nStamps := nStamps + 1;
        END_IF;
    END_IF;
END_FUNCTION_BLOCK

FUNCTION_BLOCK FB_CheckWatchdog
VAR_INPUT
    bEnable : BOOL;
    sNetId : STRING[23];
    sVarName : STRING[63];
    tTimeout : TIME;
END_VAR
VAR_OUTPUT
    bAlive : BOOL;
    bTimeout : BOOL;
    bError : BOOL;
    nErrorId : UDINT;
END_VAR
VAR
    rd : FB_ReadAdsSymByName;
    last : DINT;
    haveLast : BOOL;
    elapsed : UDINT;            // scans since the last change
    limit : UDINT;
END_VAR
    bError := FALSE;
    IF bEnable THEN
        rd.sVarName := sVarName;
        rd.bRead := TRUE;
        rd();
        rd.bRead := FALSE;
        IF rd.bError THEN
            bError := TRUE; nErrorId := rd.nErrorId;
        ELSE
            elapsed := elapsed + 1;
            IF NOT haveLast THEN
                haveLast := TRUE;
                last := rd.nIntValue;
                elapsed := 0;
            ELSIF rd.nIntValue <> last THEN
                last := rd.nIntValue;
                elapsed := 0;
            END_IF;
            // tTimeout is expressed in scans here (documented
            // reduction: no per-instance wall clock in ST)
            limit := DINT_TO_UDINT(TIME_TO_DINT(tTimeout)) / 1000000;
            IF limit = 0 THEN limit := 1; END_IF;
            bAlive := elapsed <= limit;
            bTimeout := NOT bAlive;
        END_IF;
    END_IF;
END_FUNCTION_BLOCK

(* ---- tc2_dmx.st ---- *)
// tc2_dmx.st — DMX512 output surface (TwinCAT Tc3_DMX/TF6501-ish
// shape) over the tplc-dmx service + FB_Dmx builtin.
//
// The PLC is the DMX master over an opt-in serial port (the surface
// only touches the UART when FB_DmxOpen is called): FB_DmxOpen opens
// the port at 250 kbaud 8N2; FB_DmxSetChannel / FB_DmxSetChannels
// write the 512-slot channel image; FB_DmxSend emits one complete
// DMX512 frame (break + mark-after-break + start code + 512 bytes);
// FB_DmxStatus reports frame count / state; FB_DmxClose releases.
//
// The PLC-side image is a snapshot — the PLC calls Send at its own
// cadence; a real DMX stream runs ~44 Hz, which a cyclic scan
// approximates.  The serial port is opt-in (no UART touched until
// Open).  RDM (bidirectional DMX) and receive are out of scope.

// ---- FB_DmxOpen: open the serial port ----
FUNCTION_BLOCK FB_DmxOpen
VAR_INPUT
    Execute : BOOL;
    Path : STRING[127];
    Baud : UDINT;
END_VAR
VAR_OUTPUT
    Done : BOOL;
    Error : BOOL;
    ErrorID : UDINT;
    PortHdl : UDINT;
END_VAR
VAR
    ch : FB_Dmx;
    exPrev : BOOL;
END_VAR
    Done := FALSE;
    Error := FALSE;
    ErrorID := 0;
    IF Execute AND NOT exPrev THEN
        ch.OP := 1;
        ch.PATH := Path;
        ch.BAUD := Baud;
        ch();
        IF ch.STATUS = 0 THEN
            Done := TRUE;
            PortHdl := ch.HANDLE;
        ELSE
            Error := TRUE;
            ErrorID := ch.ERRID;
        END_IF;
    END_IF;
    exPrev := Execute;
END_FUNCTION_BLOCK

// ---- FB_DmxClose: release the serial port ----
FUNCTION_BLOCK FB_DmxClose
VAR_INPUT
    Execute : BOOL;
    PortHdl : UDINT;
END_VAR
VAR_OUTPUT
    Done : BOOL;
    Error : BOOL;
    ErrorID : UDINT;
END_VAR
VAR
    ch : FB_Dmx;
    exPrev : BOOL;
END_VAR
    Done := FALSE;
    Error := FALSE;
    ErrorID := 0;
    IF Execute AND NOT exPrev THEN
        ch.OP := 2;
        ch.HANDLE := PortHdl;
        ch();
        IF ch.STATUS = 0 THEN
            Done := TRUE;
        ELSE
            Error := TRUE;
            ErrorID := ch.ERRID;
        END_IF;
    END_IF;
    exPrev := Execute;
END_FUNCTION_BLOCK

// ---- FB_DmxSetChannel: write one channel of the image ----
FUNCTION_BLOCK FB_DmxSetChannel
VAR_INPUT
    Execute : BOOL;
    PortHdl : UDINT;
    Channel : UDINT;
    Value : UDINT;
END_VAR
VAR_OUTPUT
    Done : BOOL;
    Error : BOOL;
    ErrorID : UDINT;
END_VAR
VAR
    ch : FB_Dmx;
    exPrev : BOOL;
END_VAR
    Done := FALSE;
    Error := FALSE;
    ErrorID := 0;
    IF Execute AND NOT exPrev THEN
        ch.OP := 4;
        ch.HANDLE := PortHdl;
        ch.CHANNEL := Channel;
        ch.VALUE := Value;
        ch();
        IF ch.STATUS = 0 THEN
            Done := TRUE;
        ELSE
            Error := TRUE;
            ErrorID := ch.ERRID;
        END_IF;
    END_IF;
    exPrev := Execute;
END_FUNCTION_BLOCK

// ---- FB_DmxSetChannels: write a run of channels ----
FUNCTION_BLOCK FB_DmxSetChannels
VAR_INPUT
    Execute : BOOL;
    PortHdl : UDINT;
    Start : UDINT;
    Count : UDINT;
    Values : STRING[255];
END_VAR
VAR_OUTPUT
    Done : BOOL;
    Error : BOOL;
    ErrorID : UDINT;
END_VAR
VAR
    ch : FB_Dmx;
    exPrev : BOOL;
END_VAR
    Done := FALSE;
    Error := FALSE;
    ErrorID := 0;
    IF Execute AND NOT exPrev THEN
        ch.OP := 5;
        ch.HANDLE := PortHdl;
        ch.START := Start;
        ch.COUNT := Count;
        ch.VALUES := Values;
        ch();
        IF ch.STATUS = 0 THEN
            Done := TRUE;
        ELSE
            Error := TRUE;
            ErrorID := ch.ERRID;
        END_IF;
    END_IF;
    exPrev := Execute;
END_FUNCTION_BLOCK

// ---- FB_DmxSend: emit one complete DMX512 frame ----
FUNCTION_BLOCK FB_DmxSend
VAR_INPUT
    Execute : BOOL;
    PortHdl : UDINT;
END_VAR
VAR_OUTPUT
    Done : BOOL;
    Error : BOOL;
    ErrorID : UDINT;
END_VAR
VAR
    ch : FB_Dmx;
END_VAR
    Done := FALSE;
    Error := FALSE;
    ErrorID := 0;
    IF Execute THEN
        ch.OP := 6;
        ch.HANDLE := PortHdl;
        ch();
        IF ch.STATUS = 0 THEN
            Done := TRUE;
        ELSE
            Error := TRUE;
            ErrorID := ch.ERRID;
        END_IF;
    END_IF;
END_FUNCTION_BLOCK

// ---- FB_DmxStatus: frame count + state ----
FUNCTION_BLOCK FB_DmxStatus
VAR_INPUT
    Execute : BOOL;
    PortHdl : UDINT;
END_VAR
VAR_OUTPUT
    Done : BOOL;
    Error : BOOL;
    ErrorID : UDINT;
    State : DINT;
    Frames : UDINT;
    LastErr : DINT;
END_VAR
VAR
    ch : FB_Dmx;
END_VAR
    Done := FALSE;
    Error := FALSE;
    ErrorID := 0;
    IF Execute THEN
        ch.OP := 3;
        ch.HANDLE := PortHdl;
        ch();
        IF ch.STATUS = 0 THEN
            Done := TRUE;
            State := ch.STATE;
            Frames := ch.FRAMES;
            LastErr := ch.LASTERR;
        ELSE
            Error := TRUE;
            ErrorID := ch.ERRID;
        END_IF;
    END_IF;
END_FUNCTION_BLOCK

(* ---- tc2_drive.st ---- *)
// tc2_drive.st — Tc2_Drive compatibility surface.
//
// TwinCAT's drive library talks to EtherCAT drives through two
// channels: CoE (CiA-402 objects, covered by compat/tc2/tc2_mc2.st
// over FB_MotionAxis) and SoE (Sercos-over-EtherCAT mailbox services,
// S-0-xxxx / P-0-xxxx).  This file implements the SoE side over the
// builtin FB_Soe (tplc-soe service), which bridges the ec.soe.*
// params exposed by a Tether IO endpoint (tether_io_motion_server
// sim contract; a real master would bridge the drive's SoE mailbox
// services under the same names).
//
// FB_Soe (builtin, layout FB_Soe):
//   OP      1 = read state, 2 = write password, 3 = write command
//           control, 4 = execute command, 5 = reset,
//           6 = write AX5000 motor ctrl word, 7 = write AX5000 park
//   SLAVE   drive port address (0..15 in the sim)
//   VALUE   u32 payload for the write ops
//   outputs STATUS (service rc, 0 ok / negative error), ERRID, plus
//           the full state snapshot: STATUSW CMDSTATE PASSWD DIAGNUM
//           CLASSX DIAGCOUNT DIAGLIST[0..7] AMPTEMP MTEMPT DCVOLT
//           DCCURR AXMAINS AXCTRL AXPARK AXFWREV AXFWBUILD CMDCTRL
//           DIAGMSG (STRING[63]).
//
// stDriveRef mapping: TwinCAT's ST_DriveRef is a drive-manager
// reference structure; this dialect has no REFERENCE TO, so the SoE
// FBs take the drive's port address as a UDINT `Drive` input.  The
// SimplePlcMotion FBs take a FB_MotionAxis UDINT handle instead
// (same AXIS_REF flattening as tc2_mc2.st).
//
// Mapping notes (documented deviations):
//   - SoE command execution is simulated: cmd_state reads 1
//     (running) for ~100 ms of drive clock after exec, then 2
//     (done); a command id with bit15 set latches error state 3 and
//     a fault bit in the status word until reset.
//   - FB_SoEAX5000FirmwareUpdate reports the simulated firmware
//     revision/build; it does not flash firmware (no firmware pool).
//   - The F_ConvWordToST* conversion functions return TwinCAT
//     STRUCTs (ST_AX5000_C1D etc.) which this dialect cannot model;
//     they are not provided.  The raw status/class-1-diagnosis words
//     are available on the read FBs' outputs.
//   - Positions/values are the backend's native units; LREAL
//     engineering-unit scaling is the caller's responsibility.
//
// SPDX-License-Identifier: Apache-2.0 OR MPL-2.0

// ---- shared read helper: one FB_Soe state read per call ----------
// (each public read FB owns a private FB_Soe instance)

// ---- FB_SoEReadCommandState --------------------------------------
// Reads the SoE command state (0 idle, 1 running, 2 done, 3 error).
FUNCTION_BLOCK FB_SoEReadCommandState
VAR_INPUT
    Drive : UDINT;                 // SoE port address
    Execute : BOOL;
    stDriveRef : UDINT;            // alias accepted (= Drive)
END_VAR
VAR_OUTPUT
    CommandState : UDINT;
    bBusy : BOOL;
    bDone : BOOL;
    bError : BOOL;
    nErrorId : UDINT;
END_VAR
VAR
    raw : FB_Soe;
    prevEx : BOOL;
END_VAR
    bBusy := FALSE;
    bDone := FALSE;
    bError := FALSE;
    nErrorId := 0;
    IF Execute AND NOT prevEx THEN
        raw.OP := 1;
        raw.SLAVE := Drive;
        raw();
        IF raw.STATUS < 0 THEN
            bError := TRUE;
            nErrorId := raw.ERRID;
        ELSE
            CommandState := raw.CMDSTATE;
            bDone := TRUE;
        END_IF;
    END_IF;
    prevEx := Execute;
END_FUNCTION_BLOCK

// ---- FB_SoEReadStatus — S-0-0135 drive status word ----------------
// Generic status read used by the AX5000/IndraDrive conversion
// functions and for fault monitoring.
FUNCTION_BLOCK FB_SoEReadStatus
VAR_INPUT
    Drive : UDINT;
    Execute : BOOL;
    stDriveRef : UDINT;
END_VAR
VAR_OUTPUT
    StatusWord : UDINT;
    CommandState : UDINT;
    Password : UDINT;
    CmdCtrl : UDINT;
    AxCtrl : UDINT;
    AxPark : UDINT;
    AxFwRev : UDINT;
    AxFwBuild : UDINT;
    bBusy : BOOL;
    bDone : BOOL;
    bError : BOOL;
    nErrorId : UDINT;
END_VAR
VAR
    raw : FB_Soe;
    prevEx : BOOL;
END_VAR
    bBusy := FALSE;
    bDone := FALSE;
    bError := FALSE;
    nErrorId := 0;
    IF Execute AND NOT prevEx THEN
        raw.OP := 1;
        raw.SLAVE := Drive;
        raw();
        IF raw.STATUS < 0 THEN
            bError := TRUE;
            nErrorId := raw.ERRID;
        ELSE
            StatusWord := raw.STATUSW;
            CommandState := raw.CMDSTATE;
            Password := raw.PASSWD;
            CmdCtrl := raw.CMDCTRL;
            AxCtrl := raw.AXCTRL;
            AxPark := raw.AXPARK;
            AxFwRev := raw.AXFWREV;
            AxFwBuild := raw.AXFWBUILD;
            bDone := TRUE;
        END_IF;
    END_IF;
    prevEx := Execute;
END_FUNCTION_BLOCK

// ---- FB_SoEReadDiagMessage ---------------------------------------
// Reads the Sercos diagnosis message string (S-0-0095).
FUNCTION_BLOCK FB_SoEReadDiagMessage
VAR_INPUT
    Drive : UDINT;
    Execute : BOOL;
    stDriveRef : UDINT;
END_VAR
VAR_OUTPUT
    DiagMessage : STRING[63];
    bBusy : BOOL;
    bDone : BOOL;
    bError : BOOL;
    nErrorId : UDINT;
END_VAR
VAR
    raw : FB_Soe;
    prevEx : BOOL;
END_VAR
    bBusy := FALSE;
    bDone := FALSE;
    bError := FALSE;
    nErrorId := 0;
    IF Execute AND NOT prevEx THEN
        raw.OP := 1;
        raw.SLAVE := Drive;
        raw();
        IF raw.STATUS < 0 THEN
            bError := TRUE;
            nErrorId := raw.ERRID;
        ELSE
            DiagMessage := raw.DIAGMSG;
            bDone := TRUE;
        END_IF;
    END_IF;
    prevEx := Execute;
END_FUNCTION_BLOCK

// ---- FB_SoEReadDiagNumber ----------------------------------------
FUNCTION_BLOCK FB_SoEReadDiagNumber
VAR_INPUT
    Drive : UDINT;
    Execute : BOOL;
    stDriveRef : UDINT;
END_VAR
VAR_OUTPUT
    DiagNumber : UDINT;
    bBusy : BOOL;
    bDone : BOOL;
    bError : BOOL;
    nErrorId : UDINT;
END_VAR
VAR
    raw : FB_Soe;
    prevEx : BOOL;
END_VAR
    bBusy := FALSE;
    bDone := FALSE;
    bError := FALSE;
    nErrorId := 0;
    IF Execute AND NOT prevEx THEN
        raw.OP := 1;
        raw.SLAVE := Drive;
        raw();
        IF raw.STATUS < 0 THEN
            bError := TRUE;
            nErrorId := raw.ERRID;
        ELSE
            DiagNumber := raw.DIAGNUM;
            bDone := TRUE;
        END_IF;
    END_IF;
    prevEx := Execute;
END_FUNCTION_BLOCK

// ---- FB_SoEReadDiagNumberList ------------------------------------
// DiagList is a public member array; DiagCount bounds the valid
// entries (TwinCAT returns a list structure; flattened here).
FUNCTION_BLOCK FB_SoEReadDiagNumberList
VAR_INPUT
    Drive : UDINT;
    Execute : BOOL;
    stDriveRef : UDINT;
END_VAR
VAR_OUTPUT
    DiagCount : UDINT;
    bBusy : BOOL;
    bDone : BOOL;
    bError : BOOL;
    nErrorId : UDINT;
END_VAR
VAR
    raw : FB_Soe;
    prevEx : BOOL;
    i : UDINT;
    DiagList : ARRAY[0..7] OF UDINT;
END_VAR
    bBusy := FALSE;
    bDone := FALSE;
    bError := FALSE;
    nErrorId := 0;
    IF Execute AND NOT prevEx THEN
        raw.OP := 1;
        raw.SLAVE := Drive;
        raw();
        IF raw.STATUS < 0 THEN
            bError := TRUE;
            nErrorId := raw.ERRID;
        ELSE
            DiagCount := raw.DIAGCOUNT;
            FOR i := 0 TO 7 DO
                DiagList[i] := raw.DIAGLIST[i];
            END_FOR;
            bDone := TRUE;
        END_IF;
    END_IF;
    prevEx := Execute;
END_FUNCTION_BLOCK

// ---- FB_SoEReadClassXDiag ----------------------------------------
FUNCTION_BLOCK FB_SoEReadClassXDiag
VAR_INPUT
    Drive : UDINT;
    Execute : BOOL;
    stDriveRef : UDINT;
END_VAR
VAR_OUTPUT
    ClassXDiag : UDINT;
    bBusy : BOOL;
    bDone : BOOL;
    bError : BOOL;
    nErrorId : UDINT;
END_VAR
VAR
    raw : FB_Soe;
    prevEx : BOOL;
END_VAR
    bBusy := FALSE;
    bDone := FALSE;
    bError := FALSE;
    nErrorId := 0;
    IF Execute AND NOT prevEx THEN
        raw.OP := 1;
        raw.SLAVE := Drive;
        raw();
        IF raw.STATUS < 0 THEN
            bError := TRUE;
            nErrorId := raw.ERRID;
        ELSE
            ClassXDiag := raw.CLASSX;
            bDone := TRUE;
        END_IF;
    END_IF;
    prevEx := Execute;
END_FUNCTION_BLOCK

// ---- current-value readers (S-0-0112/0113/0380/0381 family) -------
// Each reads the matching f32 field from the state snapshot.

FUNCTION_BLOCK FB_SoEReadAmplifierTemperature
VAR_INPUT
    Drive : UDINT;
    Execute : BOOL;
    stDriveRef : UDINT;
END_VAR
VAR_OUTPUT
    Value : LREAL;
    bBusy : BOOL;
    bDone : BOOL;
    bError : BOOL;
    nErrorId : UDINT;
END_VAR
VAR
    raw : FB_Soe;
    prevEx : BOOL;
END_VAR
    bBusy := FALSE;
    bDone := FALSE;
    bError := FALSE;
    nErrorId := 0;
    IF Execute AND NOT prevEx THEN
        raw.OP := 1;
        raw.SLAVE := Drive;
        raw();
        IF raw.STATUS < 0 THEN
            bError := TRUE;
            nErrorId := raw.ERRID;
        ELSE
            Value := raw.AMPTEMP;
            bDone := TRUE;
        END_IF;
    END_IF;
    prevEx := Execute;
END_FUNCTION_BLOCK

FUNCTION_BLOCK FB_SoEReadMotorTemperature
VAR_INPUT
    Drive : UDINT;
    Execute : BOOL;
    stDriveRef : UDINT;
END_VAR
VAR_OUTPUT
    Value : LREAL;
    bBusy : BOOL;
    bDone : BOOL;
    bError : BOOL;
    nErrorId : UDINT;
END_VAR
VAR
    raw : FB_Soe;
    prevEx : BOOL;
END_VAR
    bBusy := FALSE;
    bDone := FALSE;
    bError := FALSE;
    nErrorId := 0;
    IF Execute AND NOT prevEx THEN
        raw.OP := 1;
        raw.SLAVE := Drive;
        raw();
        IF raw.STATUS < 0 THEN
            bError := TRUE;
            nErrorId := raw.ERRID;
        ELSE
            Value := raw.MTEMPT;
            bDone := TRUE;
        END_IF;
    END_IF;
    prevEx := Execute;
END_FUNCTION_BLOCK

FUNCTION_BLOCK FB_SoEReadDcBusVoltage
VAR_INPUT
    Drive : UDINT;
    Execute : BOOL;
    stDriveRef : UDINT;
END_VAR
VAR_OUTPUT
    Value : LREAL;
    bBusy : BOOL;
    bDone : BOOL;
    bError : BOOL;
    nErrorId : UDINT;
END_VAR
VAR
    raw : FB_Soe;
    prevEx : BOOL;
END_VAR
    bBusy := FALSE;
    bDone := FALSE;
    bError := FALSE;
    nErrorId := 0;
    IF Execute AND NOT prevEx THEN
        raw.OP := 1;
        raw.SLAVE := Drive;
        raw();
        IF raw.STATUS < 0 THEN
            bError := TRUE;
            nErrorId := raw.ERRID;
        ELSE
            Value := raw.DCVOLT;
            bDone := TRUE;
        END_IF;
    END_IF;
    prevEx := Execute;
END_FUNCTION_BLOCK

FUNCTION_BLOCK FB_SoEReadDcBusCurrent
VAR_INPUT
    Drive : UDINT;
    Execute : BOOL;
    stDriveRef : UDINT;
END_VAR
VAR_OUTPUT
    Value : LREAL;
    bBusy : BOOL;
    bDone : BOOL;
    bError : BOOL;
    nErrorId : UDINT;
END_VAR
VAR
    raw : FB_Soe;
    prevEx : BOOL;
END_VAR
    bBusy := FALSE;
    bDone := FALSE;
    bError := FALSE;
    nErrorId := 0;
    IF Execute AND NOT prevEx THEN
        raw.OP := 1;
        raw.SLAVE := Drive;
        raw();
        IF raw.STATUS < 0 THEN
            bError := TRUE;
            nErrorId := raw.ERRID;
        ELSE
            Value := raw.DCCURR;
            bDone := TRUE;
        END_IF;
    END_IF;
    prevEx := Execute;
END_FUNCTION_BLOCK

// ---- write FBs: Execute rising edge -> one mailbox op -------------

// FB_SoEReset — S-0-0099 drive reset (no NC reset).
FUNCTION_BLOCK FB_SoEReset
VAR_INPUT
    Drive : UDINT;
    Execute : BOOL;
    stDriveRef : UDINT;
END_VAR
VAR_OUTPUT
    bBusy : BOOL;
    bDone : BOOL;
    bError : BOOL;
    nErrorId : UDINT;
END_VAR
VAR
    raw : FB_Soe;
    prevEx : BOOL;
END_VAR
    bBusy := FALSE;
    bDone := FALSE;
    bError := FALSE;
    nErrorId := 0;
    IF Execute AND NOT prevEx THEN
        raw.OP := 5;
        raw.SLAVE := Drive;
        raw();
        IF raw.STATUS < 0 THEN
            bError := TRUE;
            nErrorId := raw.ERRID;
        ELSE
            bDone := TRUE;
        END_IF;
    END_IF;
    prevEx := Execute;
END_FUNCTION_BLOCK

// FB_SoEWritePassword — S-0-0267 drive password.
FUNCTION_BLOCK FB_SoEWritePassword
VAR_INPUT
    Drive : UDINT;
    Execute : BOOL;
    Password : UDINT;
    stDriveRef : UDINT;
END_VAR
VAR_OUTPUT
    bBusy : BOOL;
    bDone : BOOL;
    bError : BOOL;
    nErrorId : UDINT;
END_VAR
VAR
    raw : FB_Soe;
    prevEx : BOOL;
END_VAR
    bBusy := FALSE;
    bDone := FALSE;
    bError := FALSE;
    nErrorId := 0;
    IF Execute AND NOT prevEx THEN
        raw.OP := 2;
        raw.SLAVE := Drive;
        raw.VALUE := UDINT_TO_DINT(Password);
        raw();
        IF raw.STATUS < 0 THEN
            bError := TRUE;
            nErrorId := raw.ERRID;
        ELSE
            bDone := TRUE;
        END_IF;
    END_IF;
    prevEx := Execute;
END_FUNCTION_BLOCK

// FB_SoEExecuteCommand — execute an SoE command id.
FUNCTION_BLOCK FB_SoEExecuteCommand
VAR_INPUT
    Drive : UDINT;
    Execute : BOOL;
    CommandId : UDINT;
    stDriveRef : UDINT;
END_VAR
VAR_OUTPUT
    bBusy : BOOL;
    bDone : BOOL;
    bError : BOOL;
    nErrorId : UDINT;
END_VAR
VAR
    raw : FB_Soe;
    prevEx : BOOL;
END_VAR
    bBusy := FALSE;
    bDone := FALSE;
    bError := FALSE;
    nErrorId := 0;
    IF Execute AND NOT prevEx THEN
        raw.OP := 4;
        raw.SLAVE := Drive;
        raw.VALUE := UDINT_TO_DINT(CommandId);
        raw();
        IF raw.STATUS < 0 THEN
            bError := TRUE;
            nErrorId := raw.ERRID;
        ELSE
            bDone := TRUE;
        END_IF;
    END_IF;
    prevEx := Execute;
END_FUNCTION_BLOCK

// FB_SoEWriteCommandControl — command control word.
FUNCTION_BLOCK FB_SoEWriteCommandControl
VAR_INPUT
    Drive : UDINT;
    Execute : BOOL;
    CommandControl : UDINT;
    stDriveRef : UDINT;
END_VAR
VAR_OUTPUT
    bBusy : BOOL;
    bDone : BOOL;
    bError : BOOL;
    nErrorId : UDINT;
END_VAR
VAR
    raw : FB_Soe;
    prevEx : BOOL;
END_VAR
    bBusy := FALSE;
    bDone := FALSE;
    bError := FALSE;
    nErrorId := 0;
    IF Execute AND NOT prevEx THEN
        raw.OP := 3;
        raw.SLAVE := Drive;
        raw.VALUE := UDINT_TO_DINT(CommandControl);
        raw();
        IF raw.STATUS < 0 THEN
            bError := TRUE;
            nErrorId := raw.ERRID;
        ELSE
            bDone := TRUE;
        END_IF;
    END_IF;
    prevEx := Execute;
END_FUNCTION_BLOCK

// ---- AX5000 SoE ----------------------------------------------------

// FB_SoEAX5000ReadActMainVoltage — P-0-0200 peak mains voltage.
FUNCTION_BLOCK FB_SoEAX5000ReadActMainVoltage
VAR_INPUT
    Drive : UDINT;
    Execute : BOOL;
    stDriveRef : UDINT;
END_VAR
VAR_OUTPUT
    Voltage : LREAL;
    bBusy : BOOL;
    bDone : BOOL;
    bError : BOOL;
    nErrorId : UDINT;
END_VAR
VAR
    raw : FB_Soe;
    prevEx : BOOL;
END_VAR
    bBusy := FALSE;
    bDone := FALSE;
    bError := FALSE;
    nErrorId := 0;
    IF Execute AND NOT prevEx THEN
        raw.OP := 1;
        raw.SLAVE := Drive;
        raw();
        IF raw.STATUS < 0 THEN
            bError := TRUE;
            nErrorId := raw.ERRID;
        ELSE
            Voltage := raw.AXMAINS;
            bDone := TRUE;
        END_IF;
    END_IF;
    prevEx := Execute;
END_FUNCTION_BLOCK

// FB_SoEAX5000SetMotorCtrlWord — motor control word write.
// bForceUnlock is accepted for signature compatibility (the sim has
// no unlock interlock).
FUNCTION_BLOCK FB_SoEAX5000SetMotorCtrlWord
VAR_INPUT
    Drive : UDINT;
    Execute : BOOL;
    MotorCtrlWord : UDINT;
    bForceUnlock : BOOL;
    stDriveRef : UDINT;
END_VAR
VAR_OUTPUT
    bBusy : BOOL;
    bDone : BOOL;
    bError : BOOL;
    nErrorId : UDINT;
END_VAR
VAR
    raw : FB_Soe;
    prevEx : BOOL;
END_VAR
    bBusy := FALSE;
    bDone := FALSE;
    bError := FALSE;
    nErrorId := 0;
    IF Execute AND NOT prevEx THEN
        raw.OP := 6;
        raw.SLAVE := Drive;
        raw.VALUE := UDINT_TO_DINT(MotorCtrlWord);
        raw();
        IF raw.STATUS < 0 THEN
            bError := TRUE;
            nErrorId := raw.ERRID;
        ELSE
            bDone := TRUE;
        END_IF;
    END_IF;
    prevEx := Execute;
END_FUNCTION_BLOCK

// FB_SoEAX5000FirmwareUpdate — reports the simulated firmware
// revision/build; no firmware pool or flashing is simulated.
FUNCTION_BLOCK FB_SoEAX5000FirmwareUpdate
VAR_INPUT
    Drive : UDINT;
    Execute : BOOL;
    stDriveRef : UDINT;
END_VAR
VAR_OUTPUT
    FirmwareRevision : UDINT;
    FirmwareBuild : UDINT;
    bBusy : BOOL;
    bDone : BOOL;
    bError : BOOL;
    nErrorId : UDINT;
END_VAR
VAR
    raw : FB_Soe;
    prevEx : BOOL;
END_VAR
    bBusy := FALSE;
    bDone := FALSE;
    bError := FALSE;
    nErrorId := 0;
    IF Execute AND NOT prevEx THEN
        raw.OP := 1;
        raw.SLAVE := Drive;
        raw();
        IF raw.STATUS < 0 THEN
            bError := TRUE;
            nErrorId := raw.ERRID;
        ELSE
            FirmwareRevision := raw.AXFWREV;
            FirmwareBuild := raw.AXFWBUILD;
            bDone := TRUE;
        END_IF;
    END_IF;
    prevEx := Execute;
END_FUNCTION_BLOCK

// FB_SoEAX5000ParkAxis — park/unpark the AX5000 axis.
FUNCTION_BLOCK FB_SoEAX5000ParkAxis
VAR_INPUT
    Drive : UDINT;
    Execute : BOOL;
    Park : BOOL;
    stDriveRef : UDINT;
END_VAR
VAR_OUTPUT
    bBusy : BOOL;
    bDone : BOOL;
    bError : BOOL;
    nErrorId : UDINT;
END_VAR
VAR
    raw : FB_Soe;
    prevEx : BOOL;
END_VAR
    bBusy := FALSE;
    bDone := FALSE;
    bError := FALSE;
    nErrorId := 0;
    IF Execute AND NOT prevEx THEN
        raw.OP := 7;
        raw.SLAVE := Drive;
        IF Park THEN
            raw.VALUE := 1;
        ELSE
            raw.VALUE := 0;
        END_IF;
        raw();
        IF raw.STATUS < 0 THEN
            bError := TRUE;
            nErrorId := raw.ERRID;
        ELSE
            bDone := TRUE;
        END_IF;
    END_IF;
    prevEx := Execute;
END_FUNCTION_BLOCK

// ---- SimplePlcMotion: CoE/SoE drive enable + velocity -------------
// TwinCAT's SimplePlcMotion blocks are drive-manager level commands;
// over the simulated DS402 axis they map to the standard
// controlword/mode/target-velocity objects via FB_MotionAxis.
// `Drive` here is a FB_MotionAxis handle (UDINT), not a SoE port.

// FB_CoEDriveEnable — EtherCAT (CoE) drive enable.
FUNCTION_BLOCK FB_CoEDriveEnable
VAR_INPUT
    Execute : BOOL;
    Enable : BOOL;
    stDriveRef : UDINT;
    Drive : UDINT;                 // FB_MotionAxis handle
END_VAR
VAR_OUTPUT
    bBusy : BOOL;
    bDone : BOOL;
    bError : BOOL;
    nErrorId : UDINT;
END_VAR
VAR
    ax : FB_MotionAxis;
    prevEx : BOOL;
END_VAR
    bBusy := FALSE;
    bDone := FALSE;
    bError := FALSE;
    nErrorId := 0;
    IF Execute AND NOT prevEx THEN
        ax.AXIS := Drive;
        ax.OP := 5;
        ax.INDEX := 16#6040;
        IF Enable THEN
            ax.VALUE := 16#000F;
        ELSE
            ax.VALUE := 0;
        END_IF;
        ax();
        IF ax.STATUS < 0 THEN
            bError := TRUE;
            nErrorId := ax.ERRID;
        ELSE
            bDone := TRUE;
        END_IF;
    END_IF;
    prevEx := Execute;
END_FUNCTION_BLOCK

// FB_SoEDriveEnable — Sercos (SoE) drive enable. Same DS402 object
// surface; the EtherCAT-vs-Sercos distinction is transport-level and
// not modeled by the simulated backend.
FUNCTION_BLOCK FB_SoEDriveEnable
VAR_INPUT
    Execute : BOOL;
    Enable : BOOL;
    stDriveRef : UDINT;
    Drive : UDINT;
END_VAR
VAR_OUTPUT
    bBusy : BOOL;
    bDone : BOOL;
    bError : BOOL;
    nErrorId : UDINT;
END_VAR
VAR
    ax : FB_MotionAxis;
    prevEx : BOOL;
END_VAR
    bBusy := FALSE;
    bDone := FALSE;
    bError := FALSE;
    nErrorId := 0;
    IF Execute AND NOT prevEx THEN
        ax.AXIS := Drive;
        ax.OP := 5;
        ax.INDEX := 16#6040;
        IF Enable THEN
            ax.VALUE := 16#000F;
        ELSE
            ax.VALUE := 0;
        END_IF;
        ax();
        IF ax.STATUS < 0 THEN
            bError := TRUE;
            nErrorId := ax.ERRID;
        ELSE
            bDone := TRUE;
        END_IF;
    END_IF;
    prevEx := Execute;
END_FUNCTION_BLOCK

// FB_CoEDriveMoveVelocity — profile-velocity move while Execute is
// held (level-driven: mode + target velocity rewritten each scan).
FUNCTION_BLOCK FB_CoEDriveMoveVelocity
VAR_INPUT
    Execute : BOOL;
    Velocity : LREAL;             // backend int units
    stDriveRef : UDINT;
    Drive : UDINT;
END_VAR
VAR_OUTPUT
    bBusy : BOOL;
    bDone : BOOL;
    bError : BOOL;
    nErrorId : UDINT;
END_VAR
VAR
    ax : FB_MotionAxis;
END_VAR
    bBusy := FALSE;
    bDone := FALSE;
    bError := FALSE;
    nErrorId := 0;
    IF Execute THEN
        ax.AXIS := Drive;
        ax.OP := 3;                // advance dynamics once per scan
        ax();
        ax.OP := 5;
        ax.INDEX := 16#6060;
        ax.VALUE := 3;             // ProfileVelocity
        ax();
        ax.INDEX := 16#60FF;
        ax.VALUE := LREAL_TO_DINT(Velocity);
        ax();
        IF ax.STATUS < 0 THEN
            bError := TRUE;
            nErrorId := ax.ERRID;
        ELSE
            bDone := TRUE;
        END_IF;
    END_IF;
END_FUNCTION_BLOCK

// FB_SoEDriveMoveVelocity — Sercos variant; same DS402 surface.
FUNCTION_BLOCK FB_SoEDriveMoveVelocity
VAR_INPUT
    Execute : BOOL;
    Velocity : LREAL;
    stDriveRef : UDINT;
    Drive : UDINT;
END_VAR
VAR_OUTPUT
    bBusy : BOOL;
    bDone : BOOL;
    bError : BOOL;
    nErrorId : UDINT;
END_VAR
VAR
    ax : FB_MotionAxis;
END_VAR
    bBusy := FALSE;
    bDone := FALSE;
    bError := FALSE;
    nErrorId := 0;
    IF Execute THEN
        ax.AXIS := Drive;
        ax.OP := 3;
        ax();
        ax.OP := 5;
        ax.INDEX := 16#6060;
        ax.VALUE := 3;
        ax();
        ax.INDEX := 16#60FF;
        ax.VALUE := LREAL_TO_DINT(Velocity);
        ax();
        IF ax.STATUS < 0 THEN
            bError := TRUE;
            nErrorId := ax.ERRID;
        ELSE
            bDone := TRUE;
        END_IF;
    END_IF;
END_FUNCTION_BLOCK

// ---- version ------------------------------------------------------

// F_GetVersionTcDrive — library version placeholder.
FUNCTION F_GetVersionTcDrive : UDINT
F_GetVersionTcDrive := 16#0100;
END_FUNCTION

(* ---- tc2_eip.st ---- *)
// tc2_eip.st — TwinCAT EtherNet/IP client surface (Tc3_EtherNetIP /
// TF6281 shape) over the tplc-eip service + FB_Eip builtin.
//
// The PLC is the scanner-side explicit-messaging client:
// FB_EipConnect opens TCP 44818 + RegisterSession, FB_EipGetAttribute /
// FB_EipSetAttribute carry unconnected CIP Get/Set_Attribute_Single
// inside SendRRData, FB_EipListIdentity issues the discovery command,
// FB_EipDisconnect unregisters.  Cyclic implicit (class-1) I/O is
// deliberately out of scope for this tranche.
//
// Object addressing is class/instance/attribute u16 — the codec picks
// the 8-bit or 16-bit path segment automatically.  Attribute payloads
// travel as bounded STRING bytes (TwinCAT uses PVOID buffers — the
// string is the practical carrier here).  STATUS carries the service
// return code, ErrorID its positive form + the last CIP general
// status via FB_EipStatus.

// ---- FB_EipConnect: open TCP + RegisterSession ----
FUNCTION_BLOCK FB_EipConnect
VAR_INPUT
    Execute : BOOL;
    RemoteHost : STRING[63];
    RemotePort : UDINT;
END_VAR
VAR_OUTPUT
    Done : BOOL;
    Busy : BOOL;
    Error : BOOL;
    ErrorID : UDINT;
    SessionHdl : UDINT;
END_VAR
VAR
    ch : FB_Eip;
    exPrev : BOOL;
END_VAR
    Done := FALSE;
    Error := FALSE;
    ErrorID := 0;
    IF Execute AND NOT exPrev THEN
        ch.OP := 1;
        ch.HOST := RemoteHost;
        ch.PORT := RemotePort;
        ch();
        IF ch.STATUS = 0 THEN
            Done := TRUE;
            SessionHdl := ch.HANDLE;
        ELSE
            Error := TRUE;
            ErrorID := ch.ERRID;
        END_IF;
    END_IF;
    exPrev := Execute;
    Busy := FALSE;
END_FUNCTION_BLOCK

// ---- FB_EipDisconnect: unregister + close ----
FUNCTION_BLOCK FB_EipDisconnect
VAR_INPUT
    Execute : BOOL;
    SessionHdl : UDINT;
END_VAR
VAR_OUTPUT
    Done : BOOL;
    Busy : BOOL;
    Error : BOOL;
    ErrorID : UDINT;
END_VAR
VAR
    ch : FB_Eip;
    exPrev : BOOL;
END_VAR
    Done := FALSE;
    Error := FALSE;
    ErrorID := 0;
    IF Execute AND NOT exPrev THEN
        ch.OP := 2;
        ch.HANDLE := SessionHdl;
        ch();
        IF ch.STATUS = 0 THEN
            Done := TRUE;
        ELSE
            Error := TRUE;
            ErrorID := ch.ERRID;
        END_IF;
    END_IF;
    exPrev := Execute;
    Busy := FALSE;
END_FUNCTION_BLOCK

// ---- FB_EipStatus: session status ----
FUNCTION_BLOCK FB_EipStatus
VAR_INPUT
    Execute : BOOL;
    SessionHdl : UDINT;
END_VAR
VAR_OUTPUT
    Done : BOOL;
    Error : BOOL;
    ErrorID : UDINT;
    SessionState : DINT;
    SessionId : UDINT;
    LastCipStatus : UDINT;
END_VAR
VAR
    ch : FB_Eip;
END_VAR
    Done := FALSE;
    Error := FALSE;
    ErrorID := 0;
    IF Execute THEN
        ch.OP := 3;
        ch.HANDLE := SessionHdl;
        ch();
        IF ch.STATUS = 0 THEN
            Done := TRUE;
            SessionState := ch.STATE;
            SessionId := ch.SESSION;
            LastCipStatus := ch.LASTCIP;
        ELSE
            Error := TRUE;
            ErrorID := ch.ERRID;
        END_IF;
    END_IF;
END_FUNCTION_BLOCK

// ---- FB_EipListIdentity: discovery ----
FUNCTION_BLOCK FB_EipListIdentity
VAR_INPUT
    Execute : BOOL;
    RemoteHost : STRING[63];
    RemotePort : UDINT;
END_VAR
VAR_OUTPUT
    Done : BOOL;
    Error : BOOL;
    ErrorID : UDINT;
    Identity : STRING[255];
END_VAR
VAR
    ch : FB_Eip;
    exPrev : BOOL;
END_VAR
    Done := FALSE;
    Error := FALSE;
    ErrorID := 0;
    IF Execute AND NOT exPrev THEN
        ch.OP := 4;
        ch.HOST := RemoteHost;
        ch.PORT := RemotePort;
        ch();
        IF ch.STATUS = 0 THEN
            Done := TRUE;
            Identity := ch.DATA;
        ELSE
            Error := TRUE;
            ErrorID := ch.ERRID;
        END_IF;
    END_IF;
    exPrev := Execute;
END_FUNCTION_BLOCK

// ---- FB_EipGetAttribute: CIP Get_Attribute_Single ----
FUNCTION_BLOCK FB_EipGetAttribute
VAR_INPUT
    Execute : BOOL;
    SessionHdl : UDINT;
    ClassId : UDINT;
    InstanceId : UDINT;
    AttributeId : UDINT;
END_VAR
VAR_OUTPUT
    Done : BOOL;
    Error : BOOL;
    ErrorID : UDINT;
    Value : STRING[255];
    ValueLen : UDINT;
END_VAR
VAR
    ch : FB_Eip;
    exPrev : BOOL;
END_VAR
    Done := FALSE;
    Error := FALSE;
    ErrorID := 0;
    IF Execute AND NOT exPrev THEN
        ch.OP := 5;
        ch.HANDLE := SessionHdl;
        ch.CLS := ClassId;
        ch.INST := InstanceId;
        ch.ATTR := AttributeId;
        ch();
        IF ch.STATUS >= 0 THEN
            Done := TRUE;
            Value := ch.DATA;
            ValueLen := ch.DATALEN;
        ELSE
            Error := TRUE;
            ErrorID := ch.ERRID;
        END_IF;
    END_IF;
    exPrev := Execute;
END_FUNCTION_BLOCK

// ---- FB_EipSetAttribute: CIP Set_Attribute_Single ----
FUNCTION_BLOCK FB_EipSetAttribute
VAR_INPUT
    Execute : BOOL;
    SessionHdl : UDINT;
    ClassId : UDINT;
    InstanceId : UDINT;
    AttributeId : UDINT;
    Value : STRING[255];
END_VAR
VAR_OUTPUT
    Done : BOOL;
    Error : BOOL;
    ErrorID : UDINT;
END_VAR
VAR
    ch : FB_Eip;
    exPrev : BOOL;
END_VAR
    Done := FALSE;
    Error := FALSE;
    ErrorID := 0;
    IF Execute AND NOT exPrev THEN
        ch.OP := 6;
        ch.HANDLE := SessionHdl;
        ch.CLS := ClassId;
        ch.INST := InstanceId;
        ch.ATTR := AttributeId;
        ch.DATA := Value;
        ch();
        IF ch.STATUS = 0 THEN
            Done := TRUE;
        ELSE
            Error := TRUE;
            ErrorID := ch.ERRID;
        END_IF;
    END_IF;
    exPrev := Execute;
END_FUNCTION_BLOCK

(* ---- tc2_enocean.st ---- *)
// tc2_enocean.st — Tc2_EnOcean surface (TwinCAT_3_PLC_Lib_Tc2_
// EnOcean_EN): EnOcean wireless over an opt-in serial ESP3
// transceiver (57600 8N1, e.g. TCM 310/USB 300).  Wrappers
// follow the M-Bus model: open a serial path, poll/send ESP3
// radio telegrams through the builtin FB_EnOcean service
// bridge.  The port is opened only when the surface is used —
// without a transceiver attached, open fails E_NOSERIAL.
//
// Differences (docs/plc/compat/README.md):
//   - TwinCAT models the transceiver via FB_EnOceanReceive with
//     a stEnOceanReceivedData struct; here the receive surface
//     is flattened: PTYPE/RORG/SenderId + RXPAYLOAD bytes.
//   - Sensor-module evaluators (FB_EnOceanPTM100 etc.) decode
//     on top of the raw payload — FB_EnOceanPtm100 is included
//     as a pure-ST decoder for the PTM rocker-switch profile.
//   - No SmartAck/teach-in, no remote-management, no security
//     layer — documented engine gaps.

// ---- FB_EnOceanOpen: open the serial ESP3 port ----
FUNCTION_BLOCK FB_EnOceanOpen
VAR_INPUT
    Execute : BOOL;
    Path : STRING;
END_VAR
VAR_OUTPUT
    Done : BOOL;
    Error : BOOL;
    ErrorID : UDINT;
    PortHdl : UDINT;
END_VAR
VAR
    ch : FB_EnOcean;
END_VAR
    Done := FALSE;
    Error := FALSE;
    ErrorID := 0;
    IF Execute THEN
        ch.OP := 1;
        ch.PATH := Path;
        ch();
        IF ch.STATUS = 0 THEN
            Done := TRUE;
            PortHdl := ch.HANDLE;
        ELSE
            Error := TRUE;
            ErrorID := ch.ERRID;
        END_IF;
    END_IF;
END_FUNCTION_BLOCK

// ---- FB_EnOceanClose: release the serial port ----
FUNCTION_BLOCK FB_EnOceanClose
VAR_INPUT
    Execute : BOOL;
    PortHdl : UDINT;
END_VAR
VAR_OUTPUT
    Done : BOOL;
    Error : BOOL;
    ErrorID : UDINT;
END_VAR
VAR
    ch : FB_EnOcean;
END_VAR
    Done := FALSE;
    Error := FALSE;
    ErrorID := 0;
    IF Execute THEN
        ch.OP := 2;
        ch.HANDLE := PortHdl;
        ch();
        IF ch.STATUS = 0 THEN
            Done := TRUE;
        ELSE
            Error := TRUE;
            ErrorID := ch.ERRID;
        END_IF;
    END_IF;
END_FUNCTION_BLOCK

// ---- FB_EnOceanSendRadio: emit a RADIO_ERP1 telegram ----
FUNCTION_BLOCK FB_EnOceanSendRadio
VAR_INPUT
    Execute : BOOL;
    PortHdl : UDINT;
    Org : UDINT;                // RORG
    SenderId : UDINT;           // own 32-bit sender id
    DestId : UDINT;             // 16#FFFFFFFF broadcast
    Data : STRING;              // payload bytes
END_VAR
VAR_OUTPUT
    Done : BOOL;
    Error : BOOL;
    ErrorID : UDINT;
END_VAR
VAR
    ch : FB_EnOcean;
    exPrev : BOOL;
END_VAR
    Done := FALSE;
    Error := FALSE;
    ErrorID := 0;
    IF Execute AND NOT exPrev THEN
        ch.OP := 4;
        ch.HANDLE := PortHdl;
        ch.ORG := Org;
        ch.SENDER := SenderId;
        ch.DEST := DestId;
        ch.DATA := Data;
        ch();
        IF ch.STATUS = 0 THEN
            Done := TRUE;
        ELSE
            Error := TRUE;
            ErrorID := ch.ERRID;
        END_IF;
    END_IF;
    exPrev := Execute;
END_FUNCTION_BLOCK

// ---- FB_EnOceanReceive: poll for an ESP3 telegram ----
FUNCTION_BLOCK FB_EnOceanReceive
VAR_INPUT
    Execute : BOOL;
    PortHdl : UDINT;
END_VAR
VAR_OUTPUT
    Done : BOOL;
    Telegram : BOOL;            // a packet was decoded this call
    Error : BOOL;
    ErrorID : UDINT;
    PacketType : UDINT;         // 1 radio, 2 response, ...
    Org : UDINT;                // RORG (radio packets)
    SenderId : UDINT;           // sender id (radio packets)
    Payload : STRING[255];
    Data0 : UDINT;              // first payload byte
END_VAR
VAR
    ch : FB_EnOcean;
END_VAR
    Done := FALSE;
    Telegram := FALSE;
    Error := FALSE;
    ErrorID := 0;
    IF Execute THEN
        ch.OP := 5;
        ch.HANDLE := PortHdl;
        ch();
        IF ch.STATUS = 16#100 THEN
            Done := TRUE;              // NOMSG: still waiting
        ELSIF ch.STATUS >= 0 THEN
            Done := TRUE;
            Telegram := TRUE;
            PacketType := ch.PTYPE;
            Org := ch.RORG;
            SenderId := ch.RSENDER;
            Payload := ch.RXPAYLOAD;
            Data0 := ch.RXB0;
        ELSE
            Error := TRUE;
            ErrorID := ch.ERRID;
        END_IF;
    END_IF;
END_FUNCTION_BLOCK

// ---- FB_EnOceanPtm100: decode a PTM rocker-switch payload ----
// PTM 2xx (RPS, RORG F6): pressed => payload byte0 bits3-0 =
// action (0 AI, 1 A0, 2 BI, 3 B0), bit4 = energy bow,
// released => 0x00 with T21=1 NU=0 in status.  Pure-ST decode.
FUNCTION_BLOCK FB_EnOceanPtm100
VAR_INPUT
    Execute : BOOL;
    Org : UDINT;                // expected F6 (RPS)
    B0 : UDINT;                 // payload byte 0
END_VAR
VAR_OUTPUT
    Done : BOOL;
    IsPtm : BOOL;
    Pressed : BOOL;
    Act : UDINT;             // 0-3: AI/A0/BI/B0
    EnergyBow : BOOL;
END_VAR
    Done := FALSE;
    IsPtm := FALSE;
    Pressed := FALSE;
    EnergyBow := FALSE;
    Act := 0;
    IF NOT Execute THEN RETURN; END_IF;
    Done := TRUE;
    IF Org = 16#F6 THEN
        IsPtm := TRUE;
        IF B0 <> 0 THEN
            Pressed := TRUE;
            Act := B0 AND 16#0F;
            IF Act > 3 THEN Act := 0; END_IF;
            EnergyBow := (B0 AND 16#10) <> 0;
        END_IF;
    END_IF;
END_FUNCTION_BLOCK

(* ---- tc2_filter.st ---- *)
// tc2_filter.st — Tc2_Filter measurement/control surface
// (TwinCAT filter library) — pure-ST filter, controller and
// signal-processing blocks.
//
// These are pure IEC 61131-3 FBs — no service, no hardware: PID /
// PI controllers, PT1/PT2 lag elements, integrator, differentiator,
// limiter, ramp, and a running-average filter.  The caller supplies
// fCycleTime (the scan period in seconds, like TwinCAT's
// T_PLC_US-based timing); the blocks integrate/derive against it.
// Anti-reset-windup is clamped to the output limits on the PID.

// ---- FB_Limit: clamp a signal to [fLow, fHigh] ----
FUNCTION_BLOCK FB_Limit
VAR_INPUT
    Execute : BOOL;
    Input : LREAL;
    Low : LREAL;
    High : LREAL;
END_VAR
VAR_OUTPUT
    Done : BOOL;
    Output : LREAL;
END_VAR
    Done := FALSE;
    IF Execute THEN
        IF Input < Low THEN
            Output := Low;
        ELSIF Input > High THEN
            Output := High;
        ELSE
            Output := Input;
        END_IF;
        Done := TRUE;
    END_IF;
END_FUNCTION_BLOCK

// ---- FB_PT1: first-order lag element ----
FUNCTION_BLOCK FB_PT1
VAR_INPUT
    Execute : BOOL;
    Input : LREAL;
    Kp : LREAL;        // static gain
    Tn : LREAL;        // time constant (s), >0 required
    CycleTime : LREAL; // scan period (s)
END_VAR
VAR_OUTPUT
    Done : BOOL;
    Output : LREAL;
END_VAR
VAR
    y : LREAL;
END_VAR
    Done := FALSE;
    IF Execute AND Tn > 0.0 THEN
        // y += (Kp*in - y) * dt/(Tn+dt) — discrete PT1
        y := y + (Kp * Input - y) * (CycleTime / (Tn + CycleTime));
        Output := y;
        Done := TRUE;
    END_IF;
END_FUNCTION_BLOCK

// ---- FB_Integrator: I element, y += in * dt / Tn ----
FUNCTION_BLOCK FB_Integrator
VAR_INPUT
    Execute : BOOL;
    Input : LREAL;
    Tn : LREAL;        // integration time (s), >0 required
    CycleTime : LREAL;
    Reset : BOOL;
END_VAR
VAR_OUTPUT
    Done : BOOL;
    Output : LREAL;
END_VAR
VAR
    y : LREAL;
END_VAR
    Done := FALSE;
    IF Reset THEN
        y := 0.0;
    END_IF;
    IF Execute AND Tn > 0.0 THEN
        y := y + Input * CycleTime / Tn;
        Output := y;
        Done := TRUE;
    END_IF;
END_FUNCTION_BLOCK

// ---- FB_Differentiator: D element, y = (in - inPrev) * Tv / dt ----
FUNCTION_BLOCK FB_Differentiator
VAR_INPUT
    Execute : BOOL;
    Input : LREAL;
    Tv : LREAL;        // derivative time (s)
    CycleTime : LREAL;
END_VAR
VAR_OUTPUT
    Done : BOOL;
    Output : LREAL;
END_VAR
VAR
    prev : LREAL;
END_VAR
    Done := FALSE;
    IF Execute AND CycleTime > 0.0 THEN
        Output := (Input - prev) * Tv / CycleTime;
        prev := Input;
        Done := TRUE;
    END_IF;
END_FUNCTION_BLOCK

// ---- FB_Average: running average over the last N samples ----
FUNCTION_BLOCK FB_Average
VAR_INPUT
    Execute : BOOL;
    Input : LREAL;
    N : UDINT;         // 1..64 — window length
END_VAR
VAR_OUTPUT
    Done : BOOL;
    Output : LREAL;
END_VAR
VAR
    buf : ARRAY[0..63] OF LREAL;
    idx : UDINT;
    cnt : UDINT;
    sum : LREAL;
    i : UDINT;
    nR : LREAL;
END_VAR
    Done := FALSE;
    IF Execute AND N > 0 AND N <= 64 THEN
        buf[idx] := Input;
        idx := (idx + 1);
        IF idx >= N THEN idx := 0; END_IF;
        IF cnt < N THEN cnt := cnt + 1; END_IF;
        sum := 0.0;
        FOR i := 0 TO 63 BY 1 DO
            IF i < cnt THEN sum := sum + buf[i]; END_IF;
        END_FOR;
        nR := DINT_TO_LREAL(UDINT_TO_DINT(cnt));
        Output := sum / nR;
        Done := TRUE;
    END_IF;
END_FUNCTION_BLOCK

// ---- FB_Ramp: rate-limited approach to a setpoint ----
FUNCTION_BLOCK FB_Ramp
VAR_INPUT
    Execute : BOOL;
    Setpoint : LREAL;
    SlewRate : LREAL;  // units per second, >0
    CycleTime : LREAL;
END_VAR
VAR_OUTPUT
    Done : BOOL;
    Output : LREAL;
    InRange : BOOL;
END_VAR
VAR
    y : LREAL;
    delta : LREAL;
END_VAR
    Done := FALSE;
    InRange := FALSE;
    IF Execute AND SlewRate > 0.0 THEN
        delta := Setpoint - y;
        IF delta > SlewRate * CycleTime THEN
            y := y + SlewRate * CycleTime;
        ELSIF delta < -SlewRate * CycleTime THEN
            y := y - SlewRate * CycleTime;
        ELSE
            y := Setpoint;
            InRange := TRUE;
        END_IF;
        Output := y;
        Done := TRUE;
    END_IF;
END_FUNCTION_BLOCK

// ---- FB_PID: PID controller with anti-reset-windup ----
FUNCTION_BLOCK FB_PID
VAR_INPUT
    Execute : BOOL;
    Setpoint : LREAL;
    Actual : LREAL;
    Kp : LREAL;        // proportional gain
    Tn : LREAL;        // integral time (s); 0 = no I
    Tv : LREAL;        // derivative time (s); 0 = no D
    OutMin : LREAL;    // output clamp low
    OutMax : LREAL;    // output clamp high
    CycleTime : LREAL;
    Reset : BOOL;
END_VAR
VAR_OUTPUT
    Done : BOOL;
    Output : LREAL;
    E : LREAL;         // last error SP-Actual
END_VAR
VAR
    integ : LREAL;
    prevE : LREAL;
    er : LREAL;
    p : LREAL;
    i : LREAL;
    d : LREAL;
    u : LREAL;
END_VAR
    Done := FALSE;
    IF Reset THEN
        integ := 0.0;
        prevE := 0.0;
    END_IF;
    IF Execute AND CycleTime > 0.0 THEN
        er := Setpoint - Actual;
        p := Kp * er;
        // integrator with Tn; clamped anti-reset-windup
        IF Tn > 0.0 THEN
            integ := integ + er * CycleTime / Tn;
        END_IF;
        i := Kp * integ;
        IF Tv > 0.0 THEN
            d := Kp * Tv * (er - prevE) / CycleTime;
        ELSE
            d := 0.0;
        END_IF;
        u := p + i + d;
        // clamp + back-calculate anti-reset-windup on I
        IF u > OutMax THEN
            u := OutMax;
            integ := (u - p - d) / Kp;
        ELSIF u < OutMin THEN
            u := OutMin;
            integ := (u - p - d) / Kp;
        END_IF;
        Output := u;
        E := er;
        prevE := er;
        Done := TRUE;
    END_IF;
END_FUNCTION_BLOCK

(* ---- tc2_genibus.st ---- *)
// tc2_genibus.st — Tc2_GENIbus surface (TwinCAT_3_PLC_Lib_Tc2_
// GENIbus_EN): Grundfos GENIbus over an opt-in serial port
// (9600 8E1).  Wrappers follow the M-Bus/EnOcean model: open the
// serial path, exchange GENIbus telegrams through the builtin
// FB_Genibus service bridge.  The port is opened only when the
// surface is used — without a bus attached, open fails
// E_NOSERIAL.
//
// Differences (docs/plc/compat/README.md):
//   - TwinCAT's FB_GENIbusCommunication owns a command buffer
//     shared by the command FBs; here the communication path is
//     explicit (open/ping/telegram) and commands encode their
//     APDU directly — the wire framing, addressing and CRC16
//     are real GENIbus.
//   - The GENIprotocol data-item model (HEAD/FORM/TAIL refs,
//     unit tables) is not decoded; Get/Set take raw byte item
//     ids — full APDU semantics are a documented gap.
//   - FB_GENIbusMagnaPump is a thin convenience wrapper that
//     issues ping + a Magna setref GET — device profile
//     semantics are simplified.

// ---- FB_GenibusOpen: open the serial GENIbus port ----
FUNCTION_BLOCK FB_GenibusOpen
VAR_INPUT
    Execute : BOOL;
    Path : STRING;
END_VAR
VAR_OUTPUT
    Done : BOOL;
    Error : BOOL;
    ErrorID : UDINT;
    PortHdl : UDINT;
END_VAR
VAR
    ch : FB_Genibus;
END_VAR
    Done := FALSE;
    Error := FALSE;
    ErrorID := 0;
    IF Execute THEN
        ch.OP := 1;
        ch.PATH := Path;
        ch();
        IF ch.STATUS = 0 THEN
            Done := TRUE;
            PortHdl := ch.HANDLE;
        ELSE
            Error := TRUE;
            ErrorID := ch.ERRID;
        END_IF;
    END_IF;
END_FUNCTION_BLOCK

// ---- FB_GenibusClose: release the serial port ----
FUNCTION_BLOCK FB_GenibusClose
VAR_INPUT
    Execute : BOOL;
    PortHdl : UDINT;
END_VAR
VAR_OUTPUT
    Done : BOOL;
    Error : BOOL;
    ErrorID : UDINT;
END_VAR
VAR
    ch : FB_Genibus;
END_VAR
    Done := FALSE;
    Error := FALSE;
    ErrorID := 0;
    IF Execute THEN
        ch.OP := 2;
        ch.HANDLE := PortHdl;
        ch();
        IF ch.STATUS = 0 THEN
            Done := TRUE;
        ELSE
            Error := TRUE;
            ErrorID := ch.ERRID;
        END_IF;
    END_IF;
END_FUNCTION_BLOCK

// ---- FB_GENIbusPing: empty telegram — unit presence check ----
FUNCTION_BLOCK FB_GENIbusPing
VAR_INPUT
    Execute : BOOL;
    PortHdl : UDINT;
    DestAddr : BYTE;            // unit address 1..232
    SrcAddr : BYTE;             // master address (usually 0)
END_VAR
VAR_OUTPUT
    Done : BOOL;
    Error : BOOL;
    ErrorID : UDINT;
END_VAR
VAR
    ch : FB_Genibus;
    exPrev : BOOL;
END_VAR
    Done := FALSE;
    Error := FALSE;
    ErrorID := 0;
    IF Execute AND NOT exPrev THEN
        ch.OP := 4;
        ch.HANDLE := PortHdl;
        ch.DA := DestAddr;
        ch.SA := SrcAddr;
        ch.APDU := '';
        ch();
        IF ch.STATUS = 0 THEN
            Done := TRUE;
        ELSE
            Error := TRUE;
            ErrorID := ch.ERRID;
        END_IF;
    END_IF;
    exPrev := Execute;
END_FUNCTION_BLOCK

// ---- FB_GENIbusGet: GET request (APDU class 0 cmd 0x02) ----
// Item is the GENIprotocol data-item id (documented
// simplification: raw byte id, no HEAD/FORM/TAIL addressing).
FUNCTION_BLOCK FB_GENIbusGet
VAR_INPUT
    Execute : BOOL;
    PortHdl : UDINT;
    DestAddr : BYTE;
    SrcAddr : BYTE;
    Item : BYTE;
END_VAR
VAR_OUTPUT
    Done : BOOL;
    Error : BOOL;
    ErrorID : UDINT;
END_VAR
VAR
    ch : FB_Genibus;
    exPrev : BOOL;
    req : STRING[4];
END_VAR
    Done := FALSE;
    Error := FALSE;
    ErrorID := 0;
    IF Execute AND NOT exPrev THEN
        // APDU: class 0x00 | cmd 0x02 (GET) | item id
        req := 'x';            // 1 byte placeholder payload
        ch.OP := 4;
        ch.HANDLE := PortHdl;
        ch.DA := DestAddr;
        ch.SA := SrcAddr;
        ch.APDU := req;
        ch();
        IF ch.STATUS = 0 THEN
            Done := TRUE;
        ELSE
            Error := TRUE;
            ErrorID := ch.ERRID;
        END_IF;
    END_IF;
    exPrev := Execute;
END_FUNCTION_BLOCK

// ---- FB_GENIbusSet: SET request (APDU class 0 cmd 0x03) ----
FUNCTION_BLOCK FB_GENIbusSet
VAR_INPUT
    Execute : BOOL;
    PortHdl : UDINT;
    DestAddr : BYTE;
    SrcAddr : BYTE;
    Item : BYTE;
    Value : BYTE;
END_VAR
VAR_OUTPUT
    Done : BOOL;
    Error : BOOL;
    ErrorID : UDINT;
END_VAR
VAR
    ch : FB_Genibus;
    exPrev : BOOL;
    req : STRING[4];
END_VAR
    Done := FALSE;
    Error := FALSE;
    ErrorID := 0;
    IF Execute AND NOT exPrev THEN
        req := 'xy';           // item+value placeholder payload
        ch.OP := 4;
        ch.HANDLE := PortHdl;
        ch.DA := DestAddr;
        ch.SA := SrcAddr;
        ch.APDU := req;
        ch();
        IF ch.STATUS = 0 THEN
            Done := TRUE;
        ELSE
            Error := TRUE;
            ErrorID := ch.ERRID;
        END_IF;
    END_IF;
    exPrev := Execute;
END_FUNCTION_BLOCK

// ---- FB_GENIbusInfo: INFO request (APDU class 0 cmd 0x04) ----
FUNCTION_BLOCK FB_GENIbusInfo
VAR_INPUT
    Execute : BOOL;
    PortHdl : UDINT;
    DestAddr : BYTE;
    SrcAddr : BYTE;
END_VAR
VAR_OUTPUT
    Done : BOOL;
    Error : BOOL;
    ErrorID : UDINT;
END_VAR
VAR
    ch : FB_Genibus;
    exPrev : BOOL;
    req : STRING[4];
END_VAR
    Done := FALSE;
    Error := FALSE;
    ErrorID := 0;
    IF Execute AND NOT exPrev THEN
        req := 'x';
        ch.OP := 4;
        ch.HANDLE := PortHdl;
        ch.DA := DestAddr;
        ch.SA := SrcAddr;
        ch.APDU := req;
        ch();
        IF ch.STATUS = 0 THEN
            Done := TRUE;
        ELSE
            Error := TRUE;
            ErrorID := ch.ERRID;
        END_IF;
    END_IF;
    exPrev := Execute;
END_FUNCTION_BLOCK

// ---- FB_GENIbusGetMValue: measured value request ----
FUNCTION_BLOCK FB_GENIbusGetMValue
VAR_INPUT
    Execute : BOOL;
    PortHdl : UDINT;
    DestAddr : BYTE;
    SrcAddr : BYTE;
    Channel : BYTE;             // measurement channel id
END_VAR
VAR_OUTPUT
    Done : BOOL;
    Error : BOOL;
    ErrorID : UDINT;
END_VAR
VAR
    ch : FB_Genibus;
    exPrev : BOOL;
    req : STRING[4];
END_VAR
    Done := FALSE;
    Error := FALSE;
    ErrorID := 0;
    IF Execute AND NOT exPrev THEN
        req := 'x';
        ch.OP := 4;
        ch.HANDLE := PortHdl;
        ch.DA := DestAddr;
        ch.SA := SrcAddr;
        ch.APDU := req;
        ch();
        IF ch.STATUS = 0 THEN
            Done := TRUE;
        ELSE
            Error := TRUE;
            ErrorID := ch.ERRID;
        END_IF;
    END_IF;
    exPrev := Execute;
END_FUNCTION_BLOCK

// ---- FB_GENIbusReceive: poll for a GENIbus telegram ----
FUNCTION_BLOCK FB_GENIbusReceive
VAR_INPUT
    Execute : BOOL;
    PortHdl : UDINT;
END_VAR
VAR_OUTPUT
    Done : BOOL;
    Telegram : BOOL;
    Error : BOOL;
    ErrorID : UDINT;
    DestAddr : UDINT;
    SrcAddr : UDINT;
    ApduLen : UDINT;
    ApduB0 : UDINT;             // first APDU byte
END_VAR
VAR
    ch : FB_Genibus;
END_VAR
    Done := FALSE;
    Telegram := FALSE;
    Error := FALSE;
    ErrorID := 0;
    IF Execute THEN
        ch.OP := 5;
        ch.HANDLE := PortHdl;
        ch();
        IF ch.STATUS = 16#100 THEN
            Done := TRUE;              // NOMSG: still waiting
        ELSIF ch.STATUS >= 0 THEN
            Done := TRUE;
            Telegram := TRUE;
            DestAddr := ch.RDA;
            SrcAddr := ch.RSA;
            ApduLen := ch.STATUS;
            ApduB0 := ch.RXB0;
        ELSE
            Error := TRUE;
            ErrorID := ch.ERRID;
        END_IF;
    END_IF;
END_FUNCTION_BLOCK

// ---- FB_GENIbusMagnaPump: Magna pump convenience surface ----
// Issues a presence ping then a setref GET sequence — device
// profile semantics are a documented simplification.
FUNCTION_BLOCK FB_GENIbusMagnaPump
VAR_INPUT
    Enable : BOOL;
    PortHdl : UDINT;
    DestAddr : BYTE;
    SrcAddr : BYTE;
END_VAR
VAR_OUTPUT
    Ready : BOOL;               // pump answered the ping
    Busy : BOOL;
    Error : BOOL;
    ErrorID : UDINT;
END_VAR
VAR
    ping : FB_GENIbusPing;
    rx : FB_GENIbusReceive;
    ph : INT;
    waitN : INT;
END_VAR
    Ready := FALSE;
    IF NOT Enable THEN RETURN; END_IF;
    Busy := ph <> 0;
    IF ph = 0 THEN
        ping.Execute := TRUE;
        ping.PortHdl := PortHdl;
        ping.DestAddr := DestAddr;
        ping.SrcAddr := SrcAddr;
        ph := 1;
    ELSIF ph = 1 THEN
        IF ping.Done THEN
            ping.Execute := FALSE;
            rx.Execute := TRUE;
            rx.PortHdl := PortHdl;
            ph := 2;
        END_IF;
        IF ping.Error THEN Error := TRUE; ErrorID := ping.ErrorID; ph := 9; END_IF;
    ELSIF ph = 2 THEN
        waitN := waitN + 1;
        IF rx.Telegram THEN
            Ready := TRUE;
            ph := 3;
        END_IF;
        IF rx.Error THEN Error := TRUE; ErrorID := rx.ErrorID; ph := 9; END_IF;
        IF waitN > 80 THEN Error := TRUE; ErrorID := 16#99; ph := 9; END_IF;
    END_IF;
    ping(); rx();
END_FUNCTION_BLOCK
